(* IEC 61131-3 sources: plc-st-coding-agent/progress/evidence/f14_v3_parallel_20261112/jobs/custom_minimax-m27, 122 files *)

(* ---- public-easy-01.candidate_01.st ---- *)
FUNCTION_BLOCK FillingLineControl
VAR_INPUT
    bottleSensor         : BOOL;
    cleaningConfirmButton : BOOL;
    fillingConfirmButton  : BOOL;
    cappingConfirmButton  : BOOL;
    packingConfirmButton  : BOOL;
    finishedButton        : BOOL;
END_VAR

VAR_OUTPUT
    Pump_Motor      : BOOL;
    Filling_Valve   : BOOL;
    Capping_Machine : BOOL;
    Packing_Machine : BOOL;
    Completion_Light : BOOL;
END_VAR

VAR
    state : INT;
END_VAR

// State definitions:
// 0 = IDLE
// 1 = CLEANING
// 2 = FILLING
// 3 = CAPPING
// 4 = PACKAGING
// 5 = COMPLETED

// Reset all outputs at the start of each cycle
Pump_Motor      := FALSE;
Filling_Valve   := FALSE;
Capping_Machine := FALSE;
Packing_Machine := FALSE;
Completion_Light := FALSE;

CASE state OF
    0: // IDLE - Waiting for bottle
        IF bottleSensor THEN
            state := 1;
        END_IF;

    1: // CLEANING - Pump motor active
        Pump_Motor := TRUE;
        IF cleaningConfirmButton THEN
            state := 2;
        END_IF;

    2: // FILLING - Filling valve active
        Filling_Valve := TRUE;
        IF fillingConfirmButton THEN
            state := 3;
        END_IF;

    3: // CAPPING - Capping machine active
        Capping_Machine := TRUE;
        IF cappingConfirmButton THEN
            state := 4;
        END_IF;

    4: // PACKAGING - Packing machine active
        Packing_Machine := TRUE;
        IF packingConfirmButton THEN
            state := 5;
        END_IF;

    5: // COMPLETED - Completion light active
        Completion_Light := TRUE;
        IF finishedButton THEN
            state := 0;
        END_IF;

END_CASE;

END_FUNCTION_BLOCK

(* ---- public-easy-01.candidate_02.st ---- *)
FUNCTION_BLOCK FillingLineControl
VAR_INPUT
    bottleSensor          : BOOL;
    cleaningConfirmButton : BOOL;
    fillingConfirmButton  : BOOL;
    cappingConfirmButton  : BOOL;
    packingConfirmButton  : BOOL;
    finishedButton        : BOOL;
END_VAR

VAR_OUTPUT
    Pump_Motor       : BOOL;
    Filling_Valve    : BOOL;
    Capping_Machine  : BOOL;
    Packing_Machine  : BOOL;
    Completion_Light : BOOL;
END_VAR

VAR
    state : INT := 0;
END_VAR

// State: 0=IDLE, 1=CLEANING, 2=FILLING, 3=CAPPING, 4=PACKAGING, 5=COMPLETED

CASE state OF
    0: // IDLE
        IF bottleSensor THEN
            state := 1;
        END_IF;

    1: // CLEANING
        Pump_Motor := TRUE;
        IF cleaningConfirmButton THEN
            state := 2;
        END_IF;

    2: // FILLING
        Filling_Valve := TRUE;
        IF fillingConfirmButton THEN
            state := 3;
        END_IF;

    3: // CAPPING
        Capping_Machine := TRUE;
        IF cappingConfirmButton THEN
            state := 4;
        END_IF;

    4: // PACKAGING
        Packing_Machine := TRUE;
        IF packingConfirmButton THEN
            state := 5;
        END_IF;

    5: // COMPLETED
        Completion_Light := TRUE;
        IF finishedButton THEN
            state := 0;
        END_IF;

END_CASE;

END_FUNCTION_BLOCK

(* ---- public-easy-01.raw_candidate_01.st ---- *)
FUNCTION_BLOCK FillingLineControl
VAR_INPUT
    bottleSensor         : BOOL;
    cleaningConfirmButton : BOOL;
    fillingConfirmButton  : BOOL;
    cappingConfirmButton  : BOOL;
    packingConfirmButton  : BOOL;
    finishedButton        : BOOL;
END_VAR

VAR_OUTPUT
    Pump_Motor      : BOOL;
    Filling_Valve   : BOOL;
    Capping_Machine : BOOL;
    Packing_Machine : BOOL;
    Completion_Light : BOOL;
END_VAR

VAR
    state : INT;
END_VAR

// State definitions:
// 0 = IDLE
// 1 = CLEANING
// 2 = FILLING
// 3 = CAPPING
// 4 = PACKAGING
// 5 = COMPLETED

// Reset all outputs at the start of each cycle
Pump_Motor      := FALSE;
Filling_Valve   := FALSE;
Capping_Machine := FALSE;
Packing_Machine := FALSE;
Completion_Light := FALSE;

CASE state OF
    0: // IDLE - Waiting for bottle
        IF bottleSensor THEN
            state := 1;
        END_IF;

    1: // CLEANING - Pump motor active
        Pump_Motor := TRUE;
        IF cleaningConfirmButton THEN
            state := 2;
        END_IF;

    2: // FILLING - Filling valve active
        Filling_Valve := TRUE;
        IF fillingConfirmButton THEN
            state := 3;
        END_IF;

    3: // CAPPING - Capping machine active
        Capping_Machine := TRUE;
        IF cappingConfirmButton THEN
            state := 4;
        END_IF;

    4: // PACKAGING - Packing machine active
        Packing_Machine := TRUE;
        IF packingConfirmButton THEN
            state := 5;
        END_IF;

    5: // COMPLETED - Completion light active
        Completion_Light := TRUE;
        IF finishedButton THEN
            state := 0;
        END_IF;

END_CASE;

END_FUNCTION_BLOCK

(* ---- public-easy-01.raw_candidate_02.st ---- *)
FUNCTION_BLOCK FillingLineControl
VAR_INPUT
    bottleSensor          : BOOL;
    cleaningConfirmButton : BOOL;
    fillingConfirmButton  : BOOL;
    cappingConfirmButton  : BOOL;
    packingConfirmButton  : BOOL;
    finishedButton        : BOOL;
END_VAR

VAR_OUTPUT
    Pump_Motor       : BOOL;
    Filling_Valve    : BOOL;
    Capping_Machine  : BOOL;
    Packing_Machine  : BOOL;
    Completion_Light : BOOL;
END_VAR

VAR
    state : INT := 0;
END_VAR

// State: 0=IDLE, 1=CLEANING, 2=FILLING, 3=CAPPING, 4=PACKAGING, 5=COMPLETED

CASE state OF
    0: // IDLE
        IF bottleSensor THEN
            state := 1;
        END_IF;

    1: // CLEANING
        Pump_Motor := TRUE;
        IF cleaningConfirmButton THEN
            state := 2;
        END_IF;

    2: // FILLING
        Filling_Valve := TRUE;
        IF fillingConfirmButton THEN
            state := 3;
        END_IF;

    3: // CAPPING
        Capping_Machine := TRUE;
        IF cappingConfirmButton THEN
            state := 4;
        END_IF;

    4: // PACKAGING
        Packing_Machine := TRUE;
        IF packingConfirmButton THEN
            state := 5;
        END_IF;

    5: // COMPLETED
        Completion_Light := TRUE;
        IF finishedButton THEN
            state := 0;
        END_IF;

END_CASE;

END_FUNCTION_BLOCK

(* ---- public-easy-02.candidate_01.st ---- *)
FUNCTION_BLOCK FB_DualWordEdgeDetection
VAR
    prevValue : DWORD;
END_VAR

VAR_OUTPUT
    hasChanged      : BOOL := FALSE;
    hasRisingEdges  : BOOL := FALSE;
    risingBits      : DWORD := 0;
    noOfRisingBits  : USINT := 0;
    hasFallingEdges : BOOL := FALSE;
    fallingBits     : DWORD := 0;
    noOfFallingBits : USINT := 0;
END_VAR

VAR
    i : USINT;
END_VAR

risingBits  := value AND NOT prevValue;
fallingBits := NOT value AND prevValue;
hasChanged      := (value <> prevValue);
hasRisingEdges  := (risingBits <> 0);
hasFallingEdges := (fallingBits <> 0);

noOfRisingBits  := 0;
noOfFallingBits := 0;

FOR i := 0 TO 31 DO
    IF (risingBits AND SHL(DWORD#1, i)) <> 0 THEN
        noOfRisingBits := noOfRisingBits + 1;
    END_IF;
    IF (fallingBits AND SHL(DWORD#1, i)) <> 0 THEN
        noOfFallingBits := noOfFallingBits + 1;
    END_IF;
END_FOR;

prevValue := value;
END_FUNCTION_BLOCK

(* ---- public-easy-02.raw_candidate_01.st ---- *)
FUNCTION_BLOCK FB_DualWordEdgeDetection
VAR
    prevValue : DWORD;
END_VAR

VAR_OUTPUT
    hasChanged      : BOOL := FALSE;
    hasRisingEdges  : BOOL := FALSE;
    risingBits      : DWORD := 0;
    noOfRisingBits  : USINT := 0;
    hasFallingEdges : BOOL := FALSE;
    fallingBits     : DWORD := 0;
    noOfFallingBits : USINT := 0;
END_VAR

VAR
    i : USINT;
END_VAR

risingBits  := value AND NOT prevValue;
fallingBits := NOT value AND prevValue;
hasChanged      := (value <> prevValue);
hasRisingEdges  := (risingBits <> 0);
hasFallingEdges := (fallingBits <> 0);

noOfRisingBits  := 0;
noOfFallingBits := 0;

FOR i := 0 TO 31 DO
    IF (risingBits AND SHL(DWORD#1, i)) <> 0 THEN
        noOfRisingBits := noOfRisingBits + 1;
    END_IF;
    IF (fallingBits AND SHL(DWORD#1, i)) <> 0 THEN
        noOfFallingBits := noOfFallingBits + 1;
    END_IF;
END_FOR;

prevValue := value;
END_FUNCTION_BLOCK

(* ---- public-easy-03.candidate_01.st ---- *)
FUNCTION_BLOCK AlarmHysteresis
VAR_INPUT
    Value      : REAL;
    hiLevel    : REAL;
    loLevel    : REAL;
    hystWindow : REAL;
END_VAR

VAR_OUTPUT
    hiAlarm : BOOL;
    loAlarm : BOOL;
    error   : BOOL;
    status  : WORD;
END_VAR

VAR
END_VAR

error  := FALSE;
status := 16#0000;

IF loLevel >= hiLevel THEN
    error  := TRUE;
    status := 16#8001;
    RETURN;
END_IF;

IF hystWindow >= (hiLevel - loLevel) THEN
    error  := TRUE;
    status := 16#8002;
    RETURN;
END_IF;

IF Value > hiLevel THEN
    hiAlarm := TRUE;
ELSIF Value < (hiLevel - hystWindow) THEN
    hiAlarm := FALSE;
END_IF;

IF Value < loLevel THEN
    loAlarm := TRUE;
ELSIF Value > (loLevel + hystWindow) THEN
    loAlarm := FALSE;
END_IF;

END_FUNCTION_BLOCK

(* ---- public-easy-03.raw_candidate_01.st ---- *)
FUNCTION_BLOCK AlarmHysteresis
VAR_INPUT
    Value      : REAL;
    hiLevel    : REAL;
    loLevel    : REAL;
    hystWindow : REAL;
END_VAR

VAR_OUTPUT
    hiAlarm : BOOL;
    loAlarm : BOOL;
    error   : BOOL;
    status  : WORD;
END_VAR

VAR
END_VAR

error  := FALSE;
status := 16#0000;

IF loLevel >= hiLevel THEN
    error  := TRUE;
    status := 16#8001;
    RETURN;
END_IF;

IF hystWindow >= (hiLevel - loLevel) THEN
    error  := TRUE;
    status := 16#8002;
    RETURN;
END_IF;

IF Value > hiLevel THEN
    hiAlarm := TRUE;
ELSIF Value < (hiLevel - hystWindow) THEN
    hiAlarm := FALSE;
END_IF;

IF Value < loLevel THEN
    loAlarm := TRUE;
ELSIF Value > (loLevel + hystWindow) THEN
    loAlarm := FALSE;
END_IF;

END_FUNCTION_BLOCK

(* ---- public-easy-04.candidate_01.st ---- *)
FUNCTION_BLOCK JamPumpControl
VAR
    ViscosityValid : BOOL := FALSE;
    DebounceAccum  : LTIME  := LTIME#0s;
    PrevViscosity  : BOOL := FALSE;
END_VAR
VAR_OUTPUT
    VFD_RUN          : BOOL := FALSE;
    PUMP_MAINT_DUE   : BOOL := FALSE;
    PUMP_RUNTIME_ACC : LTIME  := LTIME#0s;
END_VAR
VAR_INPUT
    VISCOSITY_OK    : BOOL;
    PASTE_E_STOP_NC : BOOL;
    DebounceTime    : TIME;
    CycleTime       : TIME;
END_VAR

    // Emergency stop priority: immediate disable and clear debounce state
    IF NOT PASTE_E_STOP_NC THEN
        VFD_RUN        := FALSE;
        ViscosityValid := FALSE;
        DebounceAccum  := LTIME#0s;
        PrevViscosity  := FALSE;
        RETURN;
    END_IF;

    // Viscosity debouncing
    IF NOT VISCOSITY_OK THEN
        // Signal dropped: invalidate immediately and reset
        ViscosityValid := FALSE;
        DebounceAccum  := LTIME#0s;
        PrevViscosity  := FALSE;
    ELSE
        // Detect rising edge on VISCOSITY_OK
        IF NOT PrevViscosity THEN
            DebounceAccum := LTIME#0s;
        END_IF;

        // Accumulate debounce time for this cycle
        DebounceAccum := DebounceAccum + CycleTime;

        // Check if debounce threshold reached
        IF DebounceAccum >= DebounceTime THEN
            ViscosityValid := TRUE;
        END_IF;

        PrevViscosity := TRUE;
    END_IF;

    // Run permissive: E-stop OK AND viscosity condition valid AND signal present
    IF PASTE_E_STOP_NC AND ViscosityValid AND VISCOSITY_OK THEN
        VFD_RUN := TRUE;
    ELSE
        VFD_RUN := FALSE;
    END_IF;

    // Accumulate runtime only while pump is running
    IF VFD_RUN THEN
        PUMP_RUNTIME_ACC := PUMP_RUNTIME_ACC + CycleTime;
    END_IF;

    // Maintenance indication at 500 hours (informational, non-blocking)
    IF PUMP_RUNTIME_ACC >= T#500h THEN
        PUMP_MAINT_DUE := TRUE;
    END_IF;

END_FUNCTION_BLOCK

(* ---- public-easy-04.candidate_02.st ---- *)
FUNCTION_BLOCK JamPumpControl
VAR
    ViscosityValid : BOOL := FALSE;
    DebounceAccum  : LTIME  := LTIME#0s;
    PrevViscosity  : BOOL := FALSE;
END_VAR
VAR_OUTPUT
    VFD_RUN          : BOOL := FALSE;
    PUMP_MAINT_DUE   : BOOL := FALSE;
    PUMP_RUNTIME_ACC : LTIME  := LTIME#0s;
END_VAR
VAR_INPUT
    VISCOSITY_OK    : BOOL;
    PASTE_E_STOP_NC : BOOL;
    DebounceTime    : TIME;
    CycleTime       : TIME;
END_VAR
    // Emergency stop priority: immediate disable and clear debounce state
    IF NOT PASTE_E_STOP_NC THEN
        VFD_RUN        := FALSE;
        ViscosityValid := FALSE;
        DebounceAccum  := LTIME#0s;
        PrevViscosity  := FALSE;
        RETURN;
    END_IF;

    // Viscosity debouncing
    IF NOT VISCOSITY_OK THEN
        ViscosityValid := FALSE;
        DebounceAccum  := LTIME#0s;
        PrevViscosity  := FALSE;
    ELSE
        IF NOT PrevViscosity THEN
            DebounceAccum := LTIME#0s;
        END_IF;

        DebounceAccum := DebounceAccum + TO_LTIME(TO_ULINT(CycleTime));

        IF DebounceAccum >= TO_LTIME(TO_ULINT(DebounceTime)) THEN
            ViscosityValid := TRUE;
        END_IF;

        PrevViscosity := TRUE;
    END_IF;

    // Run permissive
    IF PASTE_E_STOP_NC AND ViscosityValid AND VISCOSITY_OK THEN
        VFD_RUN := TRUE;
    ELSE
        VFD_RUN := FALSE;
    END_IF;

    // Accumulate runtime only while pump is running
    IF VFD_RUN THEN
        PUMP_RUNTIME_ACC := PUMP_RUNTIME_ACC + TO_LTIME(TO_ULINT(CycleTime));
    END_IF;

    // Maintenance indication at 500 hours
    IF PUMP_RUNTIME_ACC >= LTIME#500h THEN
        PUMP_MAINT_DUE := TRUE;
    END_IF;

END_FUNCTION_BLOCK

(* ---- public-easy-04.raw_candidate_01.st ---- *)
FUNCTION_BLOCK JamPumpControl
VAR
    ViscosityValid : BOOL := FALSE;
    DebounceAccum  : LTIME  := LTIME#0s;
    PrevViscosity  : BOOL := FALSE;
END_VAR
VAR_OUTPUT
    VFD_RUN          : BOOL := FALSE;
    PUMP_MAINT_DUE   : BOOL := FALSE;
    PUMP_RUNTIME_ACC : LTIME  := LTIME#0s;
END_VAR
VAR_INPUT
    VISCOSITY_OK    : BOOL;
    PASTE_E_STOP_NC : BOOL;
    DebounceTime    : TIME;
    CycleTime       : TIME;
END_VAR

    // Emergency stop priority: immediate disable and clear debounce state
    IF NOT PASTE_E_STOP_NC THEN
        VFD_RUN        := FALSE;
        ViscosityValid := FALSE;
        DebounceAccum  := LTIME#0s;
        PrevViscosity  := FALSE;
        RETURN;
    END_IF;

    // Viscosity debouncing
    IF NOT VISCOSITY_OK THEN
        // Signal dropped: invalidate immediately and reset
        ViscosityValid := FALSE;
        DebounceAccum  := LTIME#0s;
        PrevViscosity  := FALSE;
    ELSE
        // Detect rising edge on VISCOSITY_OK
        IF NOT PrevViscosity THEN
            DebounceAccum := LTIME#0s;
        END_IF;

        // Accumulate debounce time for this cycle
        DebounceAccum := DebounceAccum + CycleTime;

        // Check if debounce threshold reached
        IF DebounceAccum >= DebounceTime THEN
            ViscosityValid := TRUE;
        END_IF;

        PrevViscosity := TRUE;
    END_IF;

    // Run permissive: E-stop OK AND viscosity condition valid AND signal present
    IF PASTE_E_STOP_NC AND ViscosityValid AND VISCOSITY_OK THEN
        VFD_RUN := TRUE;
    ELSE
        VFD_RUN := FALSE;
    END_IF;

    // Accumulate runtime only while pump is running
    IF VFD_RUN THEN
        PUMP_RUNTIME_ACC := PUMP_RUNTIME_ACC + CycleTime;
    END_IF;

    // Maintenance indication at 500 hours (informational, non-blocking)
    IF PUMP_RUNTIME_ACC >= T#500h THEN
        PUMP_MAINT_DUE := TRUE;
    END_IF;

END_FUNCTION_BLOCK

(* ---- public-easy-04.raw_candidate_02.st ---- *)
FUNCTION_BLOCK JamPumpControl
VAR
    ViscosityValid : BOOL := FALSE;
    DebounceAccum  : LTIME  := LTIME#0s;
    PrevViscosity  : BOOL := FALSE;
END_VAR
VAR_OUTPUT
    VFD_RUN          : BOOL := FALSE;
    PUMP_MAINT_DUE   : BOOL := FALSE;
    PUMP_RUNTIME_ACC : LTIME  := LTIME#0s;
END_VAR
VAR_INPUT
    VISCOSITY_OK    : BOOL;
    PASTE_E_STOP_NC : BOOL;
    DebounceTime    : TIME;
    CycleTime       : TIME;
END_VAR
    // Emergency stop priority: immediate disable and clear debounce state
    IF NOT PASTE_E_STOP_NC THEN
        VFD_RUN        := FALSE;
        ViscosityValid := FALSE;
        DebounceAccum  := LTIME#0s;
        PrevViscosity  := FALSE;
        RETURN;
    END_IF;

    // Viscosity debouncing
    IF NOT VISCOSITY_OK THEN
        ViscosityValid := FALSE;
        DebounceAccum  := LTIME#0s;
        PrevViscosity  := FALSE;
    ELSE
        IF NOT PrevViscosity THEN
            DebounceAccum := LTIME#0s;
        END_IF;

        DebounceAccum := DebounceAccum + TO_LTIME(TO_ULINT(CycleTime));

        IF DebounceAccum >= TO_LTIME(TO_ULINT(DebounceTime)) THEN
            ViscosityValid := TRUE;
        END_IF;

        PrevViscosity := TRUE;
    END_IF;

    // Run permissive
    IF PASTE_E_STOP_NC AND ViscosityValid AND VISCOSITY_OK THEN
        VFD_RUN := TRUE;
    ELSE
        VFD_RUN := FALSE;
    END_IF;

    // Accumulate runtime only while pump is running
    IF VFD_RUN THEN
        PUMP_RUNTIME_ACC := PUMP_RUNTIME_ACC + TO_LTIME(TO_ULINT(CycleTime));
    END_IF;

    // Maintenance indication at 500 hours
    IF PUMP_RUNTIME_ACC >= LTIME#500h THEN
        PUMP_MAINT_DUE := TRUE;
    END_IF;

END_FUNCTION_BLOCK

(* ---- public-easy-05.candidate_01.st ---- *)
FUNCTION_BLOCK Weld_Gap_Alarm
VAR_INPUT
    Gap_Exceeded    : BOOL;
    Weld_E_Stop_NC  : BOOL;
    DebounceTime    : TIME;
END_VAR
VAR_OUTPUT
    Operator_Alert        : BOOL := FALSE;
    Weld_Soft_Start_Active: BOOL := FALSE;
END_VAR
VAR
    State           : (EStop, Init, Monitor) := Init;
    Init_Timer      : TON;
    Gap_Debounce    : TON;
    Gap_Debounced   : BOOL := FALSE;
    Gap_Accumulated : LTIME := LTIME#0s;
    CycleCount      : UINT := 0;
END_VAR

// EStop has highest priority - immediate reaction before any other logic
IF NOT Weld_E_Stop_NC THEN
    Operator_Alert := FALSE;
    Weld_Soft_Start_Active := FALSE;
    Gap_Debounced := FALSE;
    Gap_Accumulated := LTIME#0s;
    Gap_Debounce(IN := FALSE);
    Gap_Debounce.PT := T#0ms;
    Init_Timer(IN := FALSE);
    Init_Timer.PT := T#0ms;
    Init_Timer.Q := FALSE;
    State := EStop;
    RETURN;
END_IF;

// EStop released - restart initialization timer
IF State = EStop THEN
    State := Init;
    Init_Timer(IN := FALSE);
END_IF;

// State machine for initialization and monitoring
CASE State OF
    Init:
        // Begin 5-second initialization inhibition
        Init_Timer(IN := TRUE, PT := T#5s);
        Weld_Soft_Start_Active := TRUE;
        Operator_Alert := FALSE;
        Gap_Debounced := FALSE;
        Gap_Accumulated := LTIME#0s;
        Gap_Debounce(IN := FALSE);
        Gap_Debounce.PT := T#0ms;

        // Transition to monitoring after initialization completes
        IF Init_Timer.Q THEN
            State := Monitor;
            Weld_Soft_Start_Active := FALSE;
        END_IF;

    Monitor:
        Init_Timer(IN := FALSE);
        Init_Timer.Q := FALSE;
        Weld_Soft_Start_Active := FALSE;

        // Gap monitoring with debounce
        IF Gap_Exceeded THEN
            // Accumulate debounce time using cycle-based increment
            Gap_Accumulated := Gap_Accumulated + TO_LTIME(CycleCount);

            // Check if debounce threshold reached
            IF Gap_Accumulated >= TO_LTIME(DebounceTime) THEN
                Gap_Debounced := TRUE;
                Operator_Alert := TRUE;
            END_IF;
        ELSE
            // Signal is FALSE - clear alarm and reset debounce
            Gap_Debounced := FALSE;
            Operator_Alert := FALSE;
            Gap_Accumulated := LTIME#0s;
        END_IF;
END_CASE;

// Track cycle time for debounce accumulation
CycleCount := TO_UINT(T#1ms) / TO_UINT(T#1ms);

END_FUNCTION_BLOCK

(* ---- public-easy-05.candidate_02.st ---- *)
TYPE GapAlarmState :
(
    EStop  := 0,
    Init   := 1,
    Monitor := 2
) END_TYPE;

FUNCTION_BLOCK Weld_Gap_Alarm
VAR_INPUT
    Gap_Exceeded   : BOOL;
    Weld_E_Stop_NC : BOOL;
    DebounceTime   : TIME;
END_VAR
VAR_OUTPUT
    Operator_Alert        : BOOL := FALSE;
    Weld_Soft_Start_Active: BOOL := FALSE;
END_VAR
VAR
    State        : GapAlarmState := Init;
    Init_Timer   : TON;
    Gap_Debounce : TON;
END_VAR

// EStop has highest priority
IF NOT Weld_E_Stop_NC THEN
    Operator_Alert        := FALSE;
    Weld_Soft_Start_Active := FALSE;
    Init_Timer(IN := FALSE);
    Gap_Debounce(IN := FALSE);
    State := EStop;
    RETURN;
END_IF;

// EStop released - transition to initialization
IF State = EStop THEN
    State := Init;
END_IF;

CASE State OF
    Init:
        Init_Timer(IN := TRUE, PT := T#5s);
        Weld_Soft_Start_Active := TRUE;
        Operator_Alert := FALSE;
        Gap_Debounce(IN := FALSE);

        IF Init_Timer.Q THEN
            State := Monitor;
            Weld_Soft_Start_Active := FALSE;
        END_IF;

    Monitor:
        Init_Timer(IN := FALSE);
        Weld_Soft_Start_Active := FALSE;

        // Debounce gap signal: timer accumulates while TRUE,
        // resets when FALSE (ET tracks elapsed time)
        Gap_Debounce(IN := Gap_Exceeded, PT := DebounceTime);

        IF Gap_Debounce.Q THEN
            Operator_Alert := TRUE;
        ELSE
            Operator_Alert := FALSE;
        END_IF;
END_CASE;

END_FUNCTION_BLOCK

(* ---- public-easy-05.raw_candidate_01.st ---- *)
FUNCTION_BLOCK Weld_Gap_Alarm
VAR_INPUT
    Gap_Exceeded    : BOOL;
    Weld_E_Stop_NC  : BOOL;
    DebounceTime    : TIME;
END_VAR
VAR_OUTPUT
    Operator_Alert        : BOOL := FALSE;
    Weld_Soft_Start_Active: BOOL := FALSE;
END_VAR
VAR
    State           : (EStop, Init, Monitor) := Init;
    Init_Timer      : TON;
    Gap_Debounce    : TON;
    Gap_Debounced   : BOOL := FALSE;
    Gap_Accumulated : LTIME := LTIME#0s;
    CycleCount      : UINT := 0;
END_VAR

// EStop has highest priority - immediate reaction before any other logic
IF NOT Weld_E_Stop_NC THEN
    Operator_Alert := FALSE;
    Weld_Soft_Start_Active := FALSE;
    Gap_Debounced := FALSE;
    Gap_Accumulated := LTIME#0s;
    Gap_Debounce(IN := FALSE);
    Gap_Debounce.PT := T#0ms;
    Init_Timer(IN := FALSE);
    Init_Timer.PT := T#0ms;
    Init_Timer.Q := FALSE;
    State := EStop;
    RETURN;
END_IF;

// EStop released - restart initialization timer
IF State = EStop THEN
    State := Init;
    Init_Timer(IN := FALSE);
END_IF;

// State machine for initialization and monitoring
CASE State OF
    Init:
        // Begin 5-second initialization inhibition
        Init_Timer(IN := TRUE, PT := T#5s);
        Weld_Soft_Start_Active := TRUE;
        Operator_Alert := FALSE;
        Gap_Debounced := FALSE;
        Gap_Accumulated := LTIME#0s;
        Gap_Debounce(IN := FALSE);
        Gap_Debounce.PT := T#0ms;

        // Transition to monitoring after initialization completes
        IF Init_Timer.Q THEN
            State := Monitor;
            Weld_Soft_Start_Active := FALSE;
        END_IF;

    Monitor:
        Init_Timer(IN := FALSE);
        Init_Timer.Q := FALSE;
        Weld_Soft_Start_Active := FALSE;

        // Gap monitoring with debounce
        IF Gap_Exceeded THEN
            // Accumulate debounce time using cycle-based increment
            Gap_Accumulated := Gap_Accumulated + TO_LTIME(CycleCount);

            // Check if debounce threshold reached
            IF Gap_Accumulated >= TO_LTIME(DebounceTime) THEN
                Gap_Debounced := TRUE;
                Operator_Alert := TRUE;
            END_IF;
        ELSE
            // Signal is FALSE - clear alarm and reset debounce
            Gap_Debounced := FALSE;
            Operator_Alert := FALSE;
            Gap_Accumulated := LTIME#0s;
        END_IF;
END_CASE;

// Track cycle time for debounce accumulation
CycleCount := TO_UINT(T#1ms) / TO_UINT(T#1ms);

END_FUNCTION_BLOCK

(* ---- public-easy-05.raw_candidate_02.st ---- *)
TYPE GapAlarmState :
(
    EStop  := 0,
    Init   := 1,
    Monitor := 2
) END_TYPE

FUNCTION_BLOCK Weld_Gap_Alarm
VAR_INPUT
    Gap_Exceeded   : BOOL;
    Weld_E_Stop_NC : BOOL;
    DebounceTime   : TIME;
END_VAR
VAR_OUTPUT
    Operator_Alert        : BOOL := FALSE;
    Weld_Soft_Start_Active: BOOL := FALSE;
END_VAR
VAR
    State        : GapAlarmState := Init;
    Init_Timer   : TON;
    Gap_Debounce : TON;
END_VAR

// EStop has highest priority
IF NOT Weld_E_Stop_NC THEN
    Operator_Alert        := FALSE;
    Weld_Soft_Start_Active := FALSE;
    Init_Timer(IN := FALSE);
    Gap_Debounce(IN := FALSE);
    State := EStop;
    RETURN;
END_IF;

// EStop released - transition to initialization
IF State = EStop THEN
    State := Init;
END_IF;

CASE State OF
    Init:
        Init_Timer(IN := TRUE, PT := T#5s);
        Weld_Soft_Start_Active := TRUE;
        Operator_Alert := FALSE;
        Gap_Debounce(IN := FALSE);

        IF Init_Timer.Q THEN
            State := Monitor;
            Weld_Soft_Start_Active := FALSE;
        END_IF;

    Monitor:
        Init_Timer(IN := FALSE);
        Weld_Soft_Start_Active := FALSE;

        // Debounce gap signal: timer accumulates while TRUE,
        // resets when FALSE (ET tracks elapsed time)
        Gap_Debounce(IN := Gap_Exceeded, PT := DebounceTime);

        IF Gap_Debounce.Q THEN
            Operator_Alert := TRUE;
        ELSE
            Operator_Alert := FALSE;
        END_IF;
END_CASE;

END_FUNCTION_BLOCK

(* ---- public-easy-06.candidate_01.st ---- *)
FUNCTION_BLOCK AerationBlowerControl
VAR_INPUT
    DO_LOW : BOOL;
    AERATION_E_STOP_NC : BOOL;
END_VAR

VAR_OUTPUT
    BLOWER_RUN : BOOL := FALSE;
    AERATION_BLOWER_CYCLE_COUNT : UINT := 0;
END_VAR

VAR
    StartDelayTimer : TON;
    BlowerRunPrev : BOOL := FALSE;
END_VAR

    // Start delay timing when both DO_LOW and E-stop inactive (NC = TRUE)
    IF DO_LOW AND AERATION_E_STOP_NC THEN
        // Start the 5-second timer
        StartDelayTimer(IN := TRUE, PT := T#5S);

        // BLOWER_RUN only TRUE after timer completes
        IF StartDelayTimer.Q THEN
            BLOWER_RUN := TRUE;
        ELSE
            BLOWER_RUN := FALSE;
        END_IF;
    ELSE
        // Conditions lost: reset timer and disable blower
        StartDelayTimer(IN := FALSE);
        BLOWER_RUN := FALSE;
    END_IF;

    // Count FALSE-to-TRUE transitions of BLOWER_RUN
    IF BLOWER_RUN AND NOT BlowerRunPrev THEN
        AERATION_BLOWER_CYCLE_COUNT := AERATION_BLOWER_CYCLE_COUNT + 1;
    END_IF;

    // Store previous state for edge detection
    BlowerRunPrev := BLOWER_RUN;

END_FUNCTION_BLOCK

(* ---- public-easy-06.raw_candidate_01.st ---- *)
FUNCTION_BLOCK AerationBlowerControl
VAR_INPUT
    DO_LOW : BOOL;
    AERATION_E_STOP_NC : BOOL;
END_VAR

VAR_OUTPUT
    BLOWER_RUN : BOOL := FALSE;
    AERATION_BLOWER_CYCLE_COUNT : UINT := 0;
END_VAR

VAR
    StartDelayTimer : TON;
    BlowerRunPrev : BOOL := FALSE;
END_VAR

    // Start delay timing when both DO_LOW and E-stop inactive (NC = TRUE)
    IF DO_LOW AND AERATION_E_STOP_NC THEN
        // Start the 5-second timer
        StartDelayTimer(IN := TRUE, PT := T#5S);

        // BLOWER_RUN only TRUE after timer completes
        IF StartDelayTimer.Q THEN
            BLOWER_RUN := TRUE;
        ELSE
            BLOWER_RUN := FALSE;
        END_IF;
    ELSE
        // Conditions lost: reset timer and disable blower
        StartDelayTimer(IN := FALSE);
        BLOWER_RUN := FALSE;
    END_IF;

    // Count FALSE-to-TRUE transitions of BLOWER_RUN
    IF BLOWER_RUN AND NOT BlowerRunPrev THEN
        AERATION_BLOWER_CYCLE_COUNT := AERATION_BLOWER_CYCLE_COUNT + 1;
    END_IF;

    // Store previous state for edge detection
    BlowerRunPrev := BLOWER_RUN;

END_FUNCTION_BLOCK

(* ---- public-hard-01.candidate_01.st ---- *)
FUNCTION_BLOCK MaterialProportioningControl
VAR_INPUT
    estop            : BOOL;
    opeMode          : BOOL;
    valveAStart      : BOOL;
    valveBStart      : BOOL;
    valveCStart      : BOOL;
    valveDStart      : BOOL;
    mixMotorStart    : BOOL;
    autoStart        : BOOL;
    processMode      : BOOL;
    levelSensor      : INT;
    mixMotorComplete : BOOL;
END_VAR
VAR_OUTPUT
    valveARun    : BOOL;
    valveBRun    : BOOL;
    valveCRun    : BOOL;
    valveDRun    : BOOL;
    mixMotorRun  : BOOL;
END_VAR
VAR
    State          : INT;
    StateNext      : INT;
    autoStarted    : BOOL;
    valveAToggled  : BOOL;
    valveBToggled  : BOOL;
    valveCToggled  : BOOL;
    valveDToggled  : BOOL;
    motorToggled   : BOOL;
    lastAutoStart  : BOOL;
    lastValveAStart : BOOL;
    lastValveBStart : BOOL;
    lastValveCStart : BOOL;
    lastValveDStart : BOOL;
    lastMixMotorStart : BOOL;
END_VAR

VAR CONSTANT
    AUTO_IDLE       : INT := 0;
    AUTO_FILL_A     : INT := 1;
    AUTO_FILL_B     : INT := 2;
    AUTO_FILL_C     : INT := 3;
    AUTO_MIXING     : INT := 4;
    AUTO_DRAIN      : INT := 5;
END_VAR

    lastAutoStart := autoStart;
    lastValveAStart := valveAStart;
    lastValveBStart := valveBStart;
    lastValveCStart := valveCStart;
    lastValveDStart := valveDStart;
    lastMixMotorStart := mixMotorStart;

    valveARun := FALSE;
    valveBRun := FALSE;
    valveCRun := FALSE;
    valveDRun := FALSE;
    mixMotorRun := FALSE;

    IF NOT estop THEN
        State := AUTO_IDLE;
        autoStarted := FALSE;
        valveAToggled := FALSE;
        valveBToggled := FALSE;
        valveCToggled := FALSE;
        valveDToggled := FALSE;
        motorToggled := FALSE;
        RETURN;
    END_IF;

    IF NOT opeMode THEN
        State := AUTO_IDLE;
        autoStarted := FALSE;

        IF valveAStart AND NOT lastValveAStart THEN
            valveAToggled := NOT valveAToggled;
        END_IF;

        IF valveBStart AND NOT lastValveBStart THEN
            valveBToggled := NOT valveBToggled;
        END_IF;

        IF valveCStart AND NOT lastValveCStart THEN
            valveCToggled := NOT valveCToggled;
        END_IF;

        IF valveDStart AND NOT lastValveDStart THEN
            valveDToggled := NOT valveDToggled;
        END_IF;

        IF mixMotorStart AND NOT lastMixMotorStart THEN
            motorToggled := NOT motorToggled;
        END_IF;

        valveARun := valveAToggled;
        valveBRun := valveBToggled;
        valveCRun := valveCToggled;
        valveDRun := valveDToggled;
        mixMotorRun := motorToggled;

        RETURN;
    END_IF;

    CASE State OF
        AUTO_IDLE:
            autoStarted := FALSE;
            valveAToggled := FALSE;
            valveBToggled := FALSE;
            valveCToggled := FALSE;
            valveDToggled := FALSE;
            motorToggled := FALSE;
            IF autoStart AND NOT lastAutoStart THEN
                State := AUTO_FILL_A;
            END_IF;

        AUTO_FILL_A:
            valveARun := TRUE;
            IF levelSensor >= 50 THEN
                valveARun := FALSE;
                State := AUTO_FILL_B;
            END_IF;

        AUTO_FILL_B:
            valveBRun := TRUE;
            IF levelSensor >= 80 THEN
                valveBRun := FALSE;
                IF NOT processMode THEN
                    State := AUTO_MIXING;
                ELSE
                    State := AUTO_FILL_C;
                END_IF;
            END_IF;

        AUTO_FILL_C:
            valveCRun := TRUE;
            IF levelSensor >= 100 THEN
                valveCRun := FALSE;
                State := AUTO_MIXING;
            END_IF;

        AUTO_MIXING:
            mixMotorRun := TRUE;
            IF mixMotorComplete THEN
                mixMotorRun := FALSE;
                State := AUTO_DRAIN;
            END_IF;

        AUTO_DRAIN:
            valveDRun := TRUE;

    END_CASE;

END_FUNCTION_BLOCK

(* ---- public-hard-01.candidate_02.st ---- *)
FUNCTION_BLOCK MaterialProportioningControl
VAR_INPUT
    estop            : BOOL;
    opeMode          : BOOL;
    valveAStart      : BOOL;
    valveBStart      : BOOL;
    valveCStart      : BOOL;
    valveDStart      : BOOL;
    mixMotorStart    : BOOL;
    autoStart        : BOOL;
    processMode      : BOOL;
    levelSensor      : INT;
    mixMotorComplete : BOOL;
END_VAR
VAR_OUTPUT
    valveARun    : BOOL;
    valveBRun    : BOOL;
    valveCRun    : BOOL;
    valveDRun    : BOOL;
    mixMotorRun  : BOOL;
END_VAR
VAR
    State             : INT;
    valveAToggled     : BOOL;
    valveBToggled     : BOOL;
    valveCToggled     : BOOL;
    valveDToggled     : BOOL;
    motorToggled      : BOOL;
    prevAutoStart     : BOOL;
    prevValveAStart   : BOOL;
    prevValveBStart   : BOOL;
    prevValveCStart   : BOOL;
    prevValveDStart   : BOOL;
    prevMixMotorStart : BOOL;
END_VAR

VAR CONSTANT
    AUTO_IDLE   : INT := 0;
    AUTO_FILL_A : INT := 1;
    AUTO_FILL_B : INT := 2;
    AUTO_FILL_C : INT := 3;
    AUTO_MIXING : INT := 4;
    AUTO_DRAIN  : INT := 5;
END_VAR

    valveARun := FALSE;
    valveBRun := FALSE;
    valveCRun := FALSE;
    valveDRun := FALSE;
    mixMotorRun := FALSE;

    IF NOT estop THEN
        State := AUTO_IDLE;
        valveAToggled := FALSE;
        valveBToggled := FALSE;
        valveCToggled := FALSE;
        valveDToggled := FALSE;
        motorToggled := FALSE;
        prevAutoStart := FALSE;
        prevValveAStart := FALSE;
        prevValveBStart := FALSE;
        prevValveCStart := FALSE;
        prevValveDStart := FALSE;
        prevMixMotorStart := FALSE;
        RETURN;
    END_IF;

    IF NOT opeMode THEN
        State := AUTO_IDLE;

        IF valveAStart AND NOT prevValveAStart THEN
            valveAToggled := NOT valveAToggled;
        END_IF;
        IF valveBStart AND NOT prevValveBStart THEN
            valveBToggled := NOT valveBToggled;
        END_IF;
        IF valveCStart AND NOT prevValveCStart THEN
            valveCToggled := NOT valveCToggled;
        END_IF;
        IF valveDStart AND NOT prevValveDStart THEN
            valveDToggled := NOT valveDToggled;
        END_IF;
        IF mixMotorStart AND NOT prevMixMotorStart THEN
            motorToggled := NOT motorToggled;
        END_IF;

        valveARun := valveAToggled;
        valveBRun := valveBToggled;
        valveCRun := valveCToggled;
        valveDRun := valveDToggled;
        mixMotorRun := motorToggled;
    ELSE
        CASE State OF
            AUTO_IDLE:
                valveAToggled := FALSE;
                valveBToggled := FALSE;
                valveCToggled := FALSE;
                valveDToggled := FALSE;
                motorToggled := FALSE;
                IF autoStart AND NOT prevAutoStart THEN
                    State := AUTO_FILL_A;
                END_IF;

            AUTO_FILL_A:
                valveARun := TRUE;
                IF levelSensor >= 50 THEN
                    valveARun := FALSE;
                    State := AUTO_FILL_B;
                END_IF;

            AUTO_FILL_B:
                valveBRun := TRUE;
                IF levelSensor >= 80 THEN
                    valveBRun := FALSE;
                    IF NOT processMode THEN
                        State := AUTO_MIXING;
                    ELSE
                        State := AUTO_FILL_C;
                    END_IF;
                END_IF;

            AUTO_FILL_C:
                valveCRun := TRUE;
                IF levelSensor >= 100 THEN
                    valveCRun := FALSE;
                    State := AUTO_MIXING;
                END_IF;

            AUTO_MIXING:
                mixMotorRun := TRUE;
                IF mixMotorComplete THEN
                    mixMotorRun := FALSE;
                    State := AUTO_DRAIN;
                END_IF;

            AUTO_DRAIN:
                valveDRun := TRUE;
        END_CASE;
    END_IF;

    prevAutoStart := autoStart;
    prevValveAStart := valveAStart;
    prevValveBStart := valveBStart;
    prevValveCStart := valveCStart;
    prevValveDStart := valveDStart;
    prevMixMotorStart := mixMotorStart;

END_FUNCTION_BLOCK

(* ---- public-hard-01.raw_candidate_01.st ---- *)
FUNCTION_BLOCK MaterialProportioningControl
VAR_INPUT
    estop            : BOOL;
    opeMode          : BOOL;
    valveAStart      : BOOL;
    valveBStart      : BOOL;
    valveCStart      : BOOL;
    valveDStart      : BOOL;
    mixMotorStart    : BOOL;
    autoStart        : BOOL;
    processMode      : BOOL;
    levelSensor      : INT;
    mixMotorComplete : BOOL;
END_VAR
VAR_OUTPUT
    valveARun    : BOOL;
    valveBRun    : BOOL;
    valveCRun    : BOOL;
    valveDRun    : BOOL;
    mixMotorRun  : BOOL;
END_VAR
VAR
    State          : INT;
    StateNext      : INT;
    autoStarted    : BOOL;
    valveAToggled  : BOOL;
    valveBToggled  : BOOL;
    valveCToggled  : BOOL;
    valveDToggled  : BOOL;
    motorToggled   : BOOL;
    lastAutoStart  : BOOL;
    lastValveAStart : BOOL;
    lastValveBStart : BOOL;
    lastValveCStart : BOOL;
    lastValveDStart : BOOL;
    lastMixMotorStart : BOOL;
END_VAR

VAR CONSTANT
    AUTO_IDLE       : INT := 0;
    AUTO_FILL_A     : INT := 1;
    AUTO_FILL_B     : INT := 2;
    AUTO_FILL_C     : INT := 3;
    AUTO_MIXING     : INT := 4;
    AUTO_DRAIN      : INT := 5;
END_VAR

    lastAutoStart := autoStart;
    lastValveAStart := valveAStart;
    lastValveBStart := valveBStart;
    lastValveCStart := valveCStart;
    lastValveDStart := valveDStart;
    lastMixMotorStart := mixMotorStart;

    valveARun := FALSE;
    valveBRun := FALSE;
    valveCRun := FALSE;
    valveDRun := FALSE;
    mixMotorRun := FALSE;

    IF NOT estop THEN
        State := AUTO_IDLE;
        autoStarted := FALSE;
        valveAToggled := FALSE;
        valveBToggled := FALSE;
        valveCToggled := FALSE;
        valveDToggled := FALSE;
        motorToggled := FALSE;
        RETURN;
    END_IF

    IF NOT opeMode THEN
        State := AUTO_IDLE;
        autoStarted := FALSE;

        IF valveAStart AND NOT lastValveAStart THEN
            valveAToggled := NOT valveAToggled;
        END_IF

        IF valveBStart AND NOT lastValveBStart THEN
            valveBToggled := NOT valveBToggled;
        END_IF

        IF valveCStart AND NOT lastValveCStart THEN
            valveCToggled := NOT valveCToggled;
        END_IF

        IF valveDStart AND NOT lastValveDStart THEN
            valveDToggled := NOT valveDToggled;
        END_IF

        IF mixMotorStart AND NOT lastMixMotorStart THEN
            motorToggled := NOT motorToggled;
        END_IF

        valveARun := valveAToggled;
        valveBRun := valveBToggled;
        valveCRun := valveCToggled;
        valveDRun := valveDToggled;
        mixMotorRun := motorToggled;

        RETURN;
    END_IF

    CASE State OF
        AUTO_IDLE:
            autoStarted := FALSE;
            valveAToggled := FALSE;
            valveBToggled := FALSE;
            valveCToggled := FALSE;
            valveDToggled := FALSE;
            motorToggled := FALSE;
            IF autoStart AND NOT lastAutoStart THEN
                State := AUTO_FILL_A;
            END_IF;

        AUTO_FILL_A:
            valveARun := TRUE;
            IF levelSensor >= 50 THEN
                valveARun := FALSE;
                State := AUTO_FILL_B;
            END_IF;

        AUTO_FILL_B:
            valveBRun := TRUE;
            IF levelSensor >= 80 THEN
                valveBRun := FALSE;
                IF NOT processMode THEN
                    State := AUTO_MIXING;
                ELSE
                    State := AUTO_FILL_C;
                END_IF;
            END_IF;

        AUTO_FILL_C:
            valveCRun := TRUE;
            IF levelSensor >= 100 THEN
                valveCRun := FALSE;
                State := AUTO_MIXING;
            END_IF;

        AUTO_MIXING:
            mixMotorRun := TRUE;
            IF mixMotorComplete THEN
                mixMotorRun := FALSE;
                State := AUTO_DRAIN;
            END_IF;

        AUTO_DRAIN:
            valveDRun := TRUE;

    END_CASE;

END_FUNCTION_BLOCK

(* ---- public-hard-01.raw_candidate_02.st ---- *)
FUNCTION_BLOCK MaterialProportioningControl
VAR_INPUT
    estop            : BOOL;
    opeMode          : BOOL;
    valveAStart      : BOOL;
    valveBStart      : BOOL;
    valveCStart      : BOOL;
    valveDStart      : BOOL;
    mixMotorStart    : BOOL;
    autoStart        : BOOL;
    processMode      : BOOL;
    levelSensor      : INT;
    mixMotorComplete : BOOL;
END_VAR
VAR_OUTPUT
    valveARun    : BOOL;
    valveBRun    : BOOL;
    valveCRun    : BOOL;
    valveDRun    : BOOL;
    mixMotorRun  : BOOL;
END_VAR
VAR
    State             : INT;
    valveAToggled     : BOOL;
    valveBToggled     : BOOL;
    valveCToggled     : BOOL;
    valveDToggled     : BOOL;
    motorToggled      : BOOL;
    prevAutoStart     : BOOL;
    prevValveAStart   : BOOL;
    prevValveBStart   : BOOL;
    prevValveCStart   : BOOL;
    prevValveDStart   : BOOL;
    prevMixMotorStart : BOOL;
END_VAR

VAR CONSTANT
    AUTO_IDLE   : INT := 0;
    AUTO_FILL_A : INT := 1;
    AUTO_FILL_B : INT := 2;
    AUTO_FILL_C : INT := 3;
    AUTO_MIXING : INT := 4;
    AUTO_DRAIN  : INT := 5;
END_VAR

    valveARun := FALSE;
    valveBRun := FALSE;
    valveCRun := FALSE;
    valveDRun := FALSE;
    mixMotorRun := FALSE;

    IF NOT estop THEN
        State := AUTO_IDLE;
        valveAToggled := FALSE;
        valveBToggled := FALSE;
        valveCToggled := FALSE;
        valveDToggled := FALSE;
        motorToggled := FALSE;
        prevAutoStart := FALSE;
        prevValveAStart := FALSE;
        prevValveBStart := FALSE;
        prevValveCStart := FALSE;
        prevValveDStart := FALSE;
        prevMixMotorStart := FALSE;
        RETURN;
    END_IF;

    IF NOT opeMode THEN
        State := AUTO_IDLE;

        IF valveAStart AND NOT prevValveAStart THEN
            valveAToggled := NOT valveAToggled;
        END_IF;
        IF valveBStart AND NOT prevValveBStart THEN
            valveBToggled := NOT valveBToggled;
        END_IF;
        IF valveCStart AND NOT prevValveCStart THEN
            valveCToggled := NOT valveCToggled;
        END_IF;
        IF valveDStart AND NOT prevValveDStart THEN
            valveDToggled := NOT valveDToggled;
        END_IF;
        IF mixMotorStart AND NOT prevMixMotorStart THEN
            motorToggled := NOT motorToggled;
        END_IF;

        valveARun := valveAToggled;
        valveBRun := valveBToggled;
        valveCRun := valveCToggled;
        valveDRun := valveDToggled;
        mixMotorRun := motorToggled;
    ELSE
        CASE State OF
            AUTO_IDLE:
                valveAToggled := FALSE;
                valveBToggled := FALSE;
                valveCToggled := FALSE;
                valveDToggled := FALSE;
                motorToggled := FALSE;
                IF autoStart AND NOT prevAutoStart THEN
                    State := AUTO_FILL_A;
                END_IF;

            AUTO_FILL_A:
                valveARun := TRUE;
                IF levelSensor >= 50 THEN
                    valveARun := FALSE;
                    State := AUTO_FILL_B;
                END_IF;

            AUTO_FILL_B:
                valveBRun := TRUE;
                IF levelSensor >= 80 THEN
                    valveBRun := FALSE;
                    IF NOT processMode THEN
                        State := AUTO_MIXING;
                    ELSE
                        State := AUTO_FILL_C;
                    END_IF;
                END_IF;

            AUTO_FILL_C:
                valveCRun := TRUE;
                IF levelSensor >= 100 THEN
                    valveCRun := FALSE;
                    State := AUTO_MIXING;
                END_IF;

            AUTO_MIXING:
                mixMotorRun := TRUE;
                IF mixMotorComplete THEN
                    mixMotorRun := FALSE;
                    State := AUTO_DRAIN;
                END_IF;

            AUTO_DRAIN:
                valveDRun := TRUE;
        END_CASE;
    END_IF;

    prevAutoStart := autoStart;
    prevValveAStart := valveAStart;
    prevValveBStart := valveBStart;
    prevValveCStart := valveCStart;
    prevValveDStart := valveDStart;
    prevMixMotorStart := mixMotorStart;

END_FUNCTION_BLOCK

(* ---- public-hard-02.candidate_01.st ---- *)
FUNCTION_BLOCK FlexibleProcessingControl
VAR_INPUT
    processLength    : USINT;
    sensor1          : BOOL;
    sensor2          : BOOL;
    sensor3          : BOOL;
    sensor4          : BOOL;
    sensor5          : BOOL;
    station1Start    : BOOL;
    station2Complete : BOOL;
    station3Complete : BOOL;
    station4Complete : BOOL;
    processSequence  : ARRAY[1..8] OF USINT;
END_VAR
VAR_OUTPUT
    conveyorLeft  : BOOL;
    conveyorRight : BOOL;
END_VAR
VAR
    state          : (STATE_IDLE, STATE_MOVING);
    currentStep    : USINT;
    targetStation  : USINT;
    currentPosition: USINT;
END_VAR

CASE state OF
STATE_IDLE:
    conveyorLeft  := FALSE;
    conveyorRight := FALSE;
    IF sensor1 AND station1Start AND processLength >= 1 THEN
        currentStep := 1;
        targetStation := processSequence[1];
        state := STATE_MOVING;
    END_IF;

STATE_MOVING:
    IF targetStation > currentPosition THEN
        conveyorRight := TRUE;
        conveyorLeft := FALSE;
        IF sensor2 AND targetStation = 2 THEN
            currentPosition := 2;
        ELSIF sensor3 AND targetStation = 3 THEN
            currentPosition := 3;
        ELSIF sensor4 AND targetStation = 4 THEN
            currentPosition := 4;
        ELSIF sensor5 AND targetStation = 5 THEN
            currentPosition := 5;
        END_IF;
    ELSIF targetStation < currentPosition THEN
        conveyorLeft  := TRUE;
        conveyorRight := FALSE;
        IF sensor4 AND targetStation = 4 THEN
            currentPosition := 4;
        ELSIF sensor3 AND targetStation = 3 THEN
            currentPosition := 3;
        ELSIF sensor2 AND targetStation = 2 THEN
            currentPosition := 2;
        ELSIF sensor1 AND targetStation = 1 THEN
            currentPosition := 1;
        END_IF;
    END_IF;
    IF currentPosition = targetStation THEN
        conveyorLeft  := FALSE;
        conveyorRight := FALSE;
        IF targetStation = 5 THEN
            state := STATE_IDLE;
        ELSE
            IF station2Complete AND targetStation = 2 THEN
                currentStep := currentStep + 1;
                IF currentStep <= processLength THEN
                    targetStation := processSequence[currentStep];
                    state := STATE_MOVING;
                ELSE
                    state := STATE_IDLE;
                END_IF;
            ELSIF station3Complete AND targetStation = 3 THEN
                currentStep := currentStep + 1;
                IF currentStep <= processLength THEN
                    targetStation := processSequence[currentStep];
                    state := STATE_MOVING;
                ELSE
                    state := STATE_IDLE;
                END_IF;
            ELSIF station4Complete AND targetStation = 4 THEN
                currentStep := currentStep + 1;
                IF currentStep <= processLength THEN
                    targetStation := processSequence[currentStep];
                    state := STATE_MOVING;
                ELSE
                    state := STATE_IDLE;
                END_IF;
            END_IF;
        END_IF;
    END_IF;
END_CASE;
END_FUNCTION_BLOCK

(* ---- public-hard-02.raw_candidate_01.st ---- *)
FUNCTION_BLOCK FlexibleProcessingControl
VAR_INPUT
    processLength    : USINT;
    sensor1          : BOOL;
    sensor2          : BOOL;
    sensor3          : BOOL;
    sensor4          : BOOL;
    sensor5          : BOOL;
    station1Start    : BOOL;
    station2Complete : BOOL;
    station3Complete : BOOL;
    station4Complete : BOOL;
    processSequence  : ARRAY[1..8] OF USINT;
END_VAR
VAR_OUTPUT
    conveyorLeft  : BOOL;
    conveyorRight : BOOL;
END_VAR
VAR
    state          : (STATE_IDLE, STATE_MOVING);
    currentStep    : USINT;
    targetStation  : USINT;
    currentPosition: USINT;
END_VAR

CASE state OF
STATE_IDLE:
    conveyorLeft  := FALSE;
    conveyorRight := FALSE;
    IF sensor1 AND station1Start AND processLength >= 1 THEN
        currentStep := 1;
        targetStation := processSequence[1];
        state := STATE_MOVING;
    END_IF

STATE_MOVING:
    IF targetStation > currentPosition THEN
        conveyorRight := TRUE;
        conveyorLeft := FALSE;
        IF sensor2 AND targetStation = 2 THEN
            currentPosition := 2;
        ELSIF sensor3 AND targetStation = 3 THEN
            currentPosition := 3;
        ELSIF sensor4 AND targetStation = 4 THEN
            currentPosition := 4;
        ELSIF sensor5 AND targetStation = 5 THEN
            currentPosition := 5;
        END_IF
    ELSIF targetStation < currentPosition THEN
        conveyorLeft  := TRUE;
        conveyorRight := FALSE;
        IF sensor4 AND targetStation = 4 THEN
            currentPosition := 4;
        ELSIF sensor3 AND targetStation = 3 THEN
            currentPosition := 3;
        ELSIF sensor2 AND targetStation = 2 THEN
            currentPosition := 2;
        ELSIF sensor1 AND targetStation = 1 THEN
            currentPosition := 1;
        END_IF
    END_IF
    IF currentPosition = targetStation THEN
        conveyorLeft  := FALSE;
        conveyorRight := FALSE;
        IF targetStation = 5 THEN
            state := STATE_IDLE;
        ELSE
            IF station2Complete AND targetStation = 2 THEN
                currentStep := currentStep + 1;
                IF currentStep <= processLength THEN
                    targetStation := processSequence[currentStep];
                    state := STATE_MOVING;
                ELSE
                    state := STATE_IDLE;
                END_IF;
            ELSIF station3Complete AND targetStation = 3 THEN
                currentStep := currentStep + 1;
                IF currentStep <= processLength THEN
                    targetStation := processSequence[currentStep];
                    state := STATE_MOVING;
                ELSE
                    state := STATE_IDLE;
                END_IF;
            ELSIF station4Complete AND targetStation = 4 THEN
                currentStep := currentStep + 1;
                IF currentStep <= processLength THEN
                    targetStation := processSequence[currentStep];
                    state := STATE_MOVING;
                ELSE
                    state := STATE_IDLE;
                END_IF;
            END_IF;
        END_IF;
    END_IF;
END_CASE;
END_FUNCTION_BLOCK

(* ---- public-hard-03.candidate_01.st ---- *)
TYPE ST_Recipe :
STRUCT
    recipeID : INT;
    ingredientType : INT;
    ingredientRatio : REAL;
    productionTemperature : REAL;
END_STRUCT;
END_TYPE;

FUNCTION_BLOCK RecipeManagement
VAR_INPUT
    addRecipe : BOOL;
    deleteRecipe : BOOL;
    modifyRecipe : BOOL;
    queryRecipe : BOOL;
    recipeIn : ST_Recipe;
END_VAR
VAR_OUTPUT
    recipeAdded : BOOL := FALSE;
    recipeDeleted : BOOL := FALSE;
    recipeModified : BOOL := FALSE;
    recipeQueryResult : ST_Recipe;
    error : BOOL := FALSE;
    status : WORD := 16#0000;
END_VAR
VAR_IN_OUT
    recipe : ARRAY[1..10] OF ST_Recipe;
END_VAR
VAR
    i : INT;
    foundIndex : INT;
    duplicateExists : BOOL;
    emptySlotIndex : INT;
END_VAR

recipeAdded := FALSE;
recipeDeleted := FALSE;
recipeModified := FALSE;
recipeQueryResult.recipeID := 0;
recipeQueryResult.ingredientType := 0;
recipeQueryResult.ingredientRatio := 0.0;
recipeQueryResult.productionTemperature := 0.0;
error := FALSE;
status := 16#0000;
foundIndex := 0;
duplicateExists := FALSE;
emptySlotIndex := 0;

IF addRecipe THEN
    duplicateExists := FALSE;
    emptySlotIndex := 0;
    FOR i := 1 TO 10 DO
        IF recipe[i].recipeID = recipeIn.recipeID AND recipeIn.recipeID <> 0 THEN
            duplicateExists := TRUE;
            EXIT;
        END_IF;
        IF recipe[i].recipeID = 0 AND emptySlotIndex = 0 THEN
            emptySlotIndex := i;
        END_IF;
    END_FOR;

    IF duplicateExists THEN
        error := TRUE;
        status := 16#8002;
    ELSIF emptySlotIndex = 0 THEN
        error := TRUE;
        status := 16#8003;
    ELSE
        recipe[emptySlotIndex].recipeID := recipeIn.recipeID;
        recipe[emptySlotIndex].ingredientType := recipeIn.ingredientType;
        recipe[emptySlotIndex].ingredientRatio := recipeIn.ingredientRatio;
        recipe[emptySlotIndex].productionTemperature := recipeIn.productionTemperature;
        recipeAdded := TRUE;
    END_IF;
END_IF;

IF deleteRecipe THEN
    foundIndex := 0;
    FOR i := 1 TO 10 DO
        IF recipe[i].recipeID = recipeIn.recipeID THEN
            foundIndex := i;
            EXIT;
        END_IF;
    END_FOR;

    IF foundIndex = 0 THEN
        error := TRUE;
        status := 16#8004;
    ELSE
        recipe[foundIndex].recipeID := 0;
        recipeDeleted := TRUE;
    END_IF;
END_IF;

IF modifyRecipe THEN
    foundIndex := 0;
    FOR i := 1 TO 10 DO
        IF recipe[i].recipeID = recipeIn.recipeID THEN
            foundIndex := i;
            EXIT;
        END_IF;
    END_FOR;

    IF foundIndex = 0 THEN
        error := TRUE;
        status := 16#8005;
    ELSE
        recipe[foundIndex].recipeID := recipeIn.recipeID;
        recipe[foundIndex].ingredientType := recipeIn.ingredientType;
        recipe[foundIndex].ingredientRatio := recipeIn.ingredientRatio;
        recipe[foundIndex].productionTemperature := recipeIn.productionTemperature;
        recipeModified := TRUE;
    END_IF;
END_IF;

IF queryRecipe THEN
    foundIndex := 0;
    FOR i := 1 TO 10 DO
        IF recipe[i].recipeID = recipeIn.recipeID THEN
            foundIndex := i;
            EXIT;
        END_IF;
    END_FOR;

    IF foundIndex = 0 THEN
        error := TRUE;
        status := 16#8001;
    ELSE
        recipeQueryResult.recipeID := recipe[foundIndex].recipeID;
        recipeQueryResult.ingredientType := recipe[foundIndex].ingredientType;
        recipeQueryResult.ingredientRatio := recipe[foundIndex].ingredientRatio;
        recipeQueryResult.productionTemperature := recipe[foundIndex].productionTemperature;
    END_IF;
END_IF;
END_FUNCTION_BLOCK

(* ---- public-hard-03.candidate_02.st ---- *)
TYPE ST_Recipe :
STRUCT
    recipeID : INT;
    ingredientType : INT;
    ingredientRatio : REAL;
    productionTemperature : REAL;
END_STRUCT;
END_TYPE;

FUNCTION_BLOCK RecipeManagement
VAR_INPUT
    addRecipe : BOOL;
    deleteRecipe : BOOL;
    modifyRecipe : BOOL;
    queryRecipe : BOOL;
    recipeIn : ST_Recipe;
END_VAR
VAR_OUTPUT
    recipeAdded : BOOL := FALSE;
    recipeDeleted : BOOL := FALSE;
    recipeModified : BOOL := FALSE;
    recipeQueryResult : ST_Recipe;
    error : BOOL := FALSE;
    status : WORD := 16#0000;
END_VAR
VAR_IN_OUT
    recipe : ARRAY[1..10] OF ST_Recipe;
END_VAR
VAR
    i : INT;
    foundIndex : INT;
    duplicateExists : BOOL;
    emptySlotIndex : INT;
END_VAR

recipeAdded := FALSE;
recipeDeleted := FALSE;
recipeModified := FALSE;
recipeQueryResult.recipeID := 0;
recipeQueryResult.ingredientType := 0;
recipeQueryResult.ingredientRatio := 0.0;
recipeQueryResult.productionTemperature := 0.0;
error := FALSE;
status := 16#0000;
foundIndex := 0;
duplicateExists := FALSE;
emptySlotIndex := 0;

IF addRecipe THEN
    duplicateExists := FALSE;
    emptySlotIndex := 0;
    FOR i := 1 TO 10 DO
        IF recipe[i].recipeID = recipeIn.recipeID AND recipeIn.recipeID <> 0 THEN
            duplicateExists := TRUE;
            EXIT;
        END_IF;
        IF recipe[i].recipeID = 0 AND emptySlotIndex = 0 THEN
            emptySlotIndex := i;
        END_IF;
    END_FOR;

    IF duplicateExists THEN
        error := TRUE;
        status := 16#8002;
    ELSIF emptySlotIndex = 0 THEN
        error := TRUE;
        status := 16#8003;
    ELSE
        recipe[emptySlotIndex].recipeID := recipeIn.recipeID;
        recipe[emptySlotIndex].ingredientType := recipeIn.ingredientType;
        recipe[emptySlotIndex].ingredientRatio := recipeIn.ingredientRatio;
        recipe[emptySlotIndex].productionTemperature := recipeIn.productionTemperature;
        recipeAdded := TRUE;
    END_IF;
END_IF;

IF deleteRecipe THEN
    foundIndex := 0;
    FOR i := 1 TO 10 DO
        IF recipe[i].recipeID = recipeIn.recipeID THEN
            foundIndex := i;
            EXIT;
        END_IF;
    END_FOR;

    IF foundIndex = 0 THEN
        error := TRUE;
        status := 16#8004;
    ELSE
        recipe[foundIndex].recipeID := 0;
        recipeDeleted := TRUE;
    END_IF;
END_IF;

IF modifyRecipe THEN
    foundIndex := 0;
    FOR i := 1 TO 10 DO
        IF recipe[i].recipeID = recipeIn.recipeID THEN
            foundIndex := i;
            EXIT;
        END_IF;
    END_FOR;

    IF foundIndex = 0 THEN
        error := TRUE;
        status := 16#8005;
    ELSE
        recipe[foundIndex].recipeID := recipeIn.recipeID;
        recipe[foundIndex].ingredientType := recipeIn.ingredientType;
        recipe[foundIndex].ingredientRatio := recipeIn.ingredientRatio;
        recipe[foundIndex].productionTemperature := recipeIn.productionTemperature;
        recipeModified := TRUE;
    END_IF;
END_IF;

IF queryRecipe THEN
    foundIndex := 0;
    FOR i := 1 TO 10 DO
        IF recipe[i].recipeID = recipeIn.recipeID THEN
            foundIndex := i;
            EXIT;
        END_IF;
    END_FOR;

    IF foundIndex = 0 THEN
        error := TRUE;
        status := 16#8001;
    ELSE
        recipeQueryResult.recipeID := recipe[foundIndex].recipeID;
        recipeQueryResult.ingredientType := recipe[foundIndex].ingredientType;
        recipeQueryResult.ingredientRatio := recipe[foundIndex].ingredientRatio;
        recipeQueryResult.productionTemperature := recipe[foundIndex].productionTemperature;
    END_IF;
END_IF;
END_FUNCTION_BLOCK

(* ---- public-hard-03.raw_candidate_01.st ---- *)
TYPE ST_Recipe :
STRUCT
    recipeID : INT;
    ingredientType : INT;
    ingredientRatio : REAL;
    productionTemperature : REAL;
END_STRUCT
END_TYPE

FUNCTION_BLOCK RecipeManagement
VAR_INPUT
    addRecipe : BOOL;
    deleteRecipe : BOOL;
    modifyRecipe : BOOL;
    queryRecipe : BOOL;
    recipeIn : ST_Recipe;
END_VAR
VAR_OUTPUT
    recipeAdded : BOOL := FALSE;
    recipeDeleted : BOOL := FALSE;
    recipeModified : BOOL := FALSE;
    recipeQueryResult : ST_Recipe;
    error : BOOL := FALSE;
    status : WORD := 16#0000;
END_VAR
VAR_IN_OUT
    recipe : ARRAY[1..10] OF ST_Recipe;
END_VAR
VAR
    i : INT;
    foundIndex : INT;
    duplicateExists : BOOL;
    emptySlotIndex : INT;
END_VAR

recipeAdded := FALSE;
recipeDeleted := FALSE;
recipeModified := FALSE;
recipeQueryResult.recipeID := 0;
recipeQueryResult.ingredientType := 0;
recipeQueryResult.ingredientRatio := 0.0;
recipeQueryResult.productionTemperature := 0.0;
error := FALSE;
status := 16#0000;
foundIndex := 0;
duplicateExists := FALSE;
emptySlotIndex := 0;

IF addRecipe THEN
    duplicateExists := FALSE;
    emptySlotIndex := 0;
    FOR i := 1 TO 10 DO
        IF recipe[i].recipeID = recipeIn.recipeID AND recipeIn.recipeID <> 0 THEN
            duplicateExists := TRUE;
            EXIT;
        END_IF
        IF recipe[i].recipeID = 0 AND emptySlotIndex = 0 THEN
            emptySlotIndex := i;
        END_IF
    END_FOR;

    IF duplicateExists THEN
        error := TRUE;
        status := 16#8002;
    ELSIF emptySlotIndex = 0 THEN
        error := TRUE;
        status := 16#8003;
    ELSE
        recipe[emptySlotIndex].recipeID := recipeIn.recipeID;
        recipe[emptySlotIndex].ingredientType := recipeIn.ingredientType;
        recipe[emptySlotIndex].ingredientRatio := recipeIn.ingredientRatio;
        recipe[emptySlotIndex].productionTemperature := recipeIn.productionTemperature;
        recipeAdded := TRUE;
    END_IF;
END_IF;

IF deleteRecipe THEN
    foundIndex := 0;
    FOR i := 1 TO 10 DO
        IF recipe[i].recipeID = recipeIn.recipeID THEN
            foundIndex := i;
            EXIT;
        END_IF
    END_FOR;

    IF foundIndex = 0 THEN
        error := TRUE;
        status := 16#8004;
    ELSE
        recipe[foundIndex].recipeID := 0;
        recipeDeleted := TRUE;
    END_IF;
END_IF;

IF modifyRecipe THEN
    foundIndex := 0;
    FOR i := 1 TO 10 DO
        IF recipe[i].recipeID = recipeIn.recipeID THEN
            foundIndex := i;
            EXIT;
        END_IF
    END_FOR;

    IF foundIndex = 0 THEN
        error := TRUE;
        status := 16#8005;
    ELSE
        recipe[foundIndex].recipeID := recipeIn.recipeID;
        recipe[foundIndex].ingredientType := recipeIn.ingredientType;
        recipe[foundIndex].ingredientRatio := recipeIn.ingredientRatio;
        recipe[foundIndex].productionTemperature := recipeIn.productionTemperature;
        recipeModified := TRUE;
    END_IF;
END_IF;

IF queryRecipe THEN
    foundIndex := 0;
    FOR i := 1 TO 10 DO
        IF recipe[i].recipeID = recipeIn.recipeID THEN
            foundIndex := i;
            EXIT;
        END_IF
    END_FOR;

    IF foundIndex = 0 THEN
        error := TRUE;
        status := 16#8001;
    ELSE
        recipeQueryResult.recipeID := recipe[foundIndex].recipeID;
        recipeQueryResult.ingredientType := recipe[foundIndex].ingredientType;
        recipeQueryResult.ingredientRatio := recipe[foundIndex].ingredientRatio;
        recipeQueryResult.productionTemperature := recipe[foundIndex].productionTemperature;
    END_IF;
END_IF;
END_FUNCTION_BLOCK

(* ---- public-hard-03.raw_candidate_02.st ---- *)
TYPE ST_Recipe :
STRUCT
    recipeID : INT;
    ingredientType : INT;
    ingredientRatio : REAL;
    productionTemperature : REAL;
END_STRUCT
END_TYPE

FUNCTION_BLOCK RecipeManagement
VAR_INPUT
    addRecipe : BOOL;
    deleteRecipe : BOOL;
    modifyRecipe : BOOL;
    queryRecipe : BOOL;
    recipeIn : ST_Recipe;
END_VAR
VAR_OUTPUT
    recipeAdded : BOOL := FALSE;
    recipeDeleted : BOOL := FALSE;
    recipeModified : BOOL := FALSE;
    recipeQueryResult : ST_Recipe;
    error : BOOL := FALSE;
    status : WORD := 16#0000;
END_VAR
VAR_IN_OUT
    recipe : ARRAY[1..10] OF ST_Recipe;
END_VAR
VAR
    i : INT;
    foundIndex : INT;
    duplicateExists : BOOL;
    emptySlotIndex : INT;
END_VAR

recipeAdded := FALSE;
recipeDeleted := FALSE;
recipeModified := FALSE;
recipeQueryResult.recipeID := 0;
recipeQueryResult.ingredientType := 0;
recipeQueryResult.ingredientRatio := 0.0;
recipeQueryResult.productionTemperature := 0.0;
error := FALSE;
status := 16#0000;
foundIndex := 0;
duplicateExists := FALSE;
emptySlotIndex := 0;

IF addRecipe THEN
    duplicateExists := FALSE;
    emptySlotIndex := 0;
    FOR i := 1 TO 10 DO
        IF recipe[i].recipeID = recipeIn.recipeID AND recipeIn.recipeID <> 0 THEN
            duplicateExists := TRUE;
            EXIT;
        END_IF;
        IF recipe[i].recipeID = 0 AND emptySlotIndex = 0 THEN
            emptySlotIndex := i;
        END_IF;
    END_FOR;

    IF duplicateExists THEN
        error := TRUE;
        status := 16#8002;
    ELSIF emptySlotIndex = 0 THEN
        error := TRUE;
        status := 16#8003;
    ELSE
        recipe[emptySlotIndex].recipeID := recipeIn.recipeID;
        recipe[emptySlotIndex].ingredientType := recipeIn.ingredientType;
        recipe[emptySlotIndex].ingredientRatio := recipeIn.ingredientRatio;
        recipe[emptySlotIndex].productionTemperature := recipeIn.productionTemperature;
        recipeAdded := TRUE;
    END_IF;
END_IF;

IF deleteRecipe THEN
    foundIndex := 0;
    FOR i := 1 TO 10 DO
        IF recipe[i].recipeID = recipeIn.recipeID THEN
            foundIndex := i;
            EXIT;
        END_IF;
    END_FOR;

    IF foundIndex = 0 THEN
        error := TRUE;
        status := 16#8004;
    ELSE
        recipe[foundIndex].recipeID := 0;
        recipeDeleted := TRUE;
    END_IF;
END_IF;

IF modifyRecipe THEN
    foundIndex := 0;
    FOR i := 1 TO 10 DO
        IF recipe[i].recipeID = recipeIn.recipeID THEN
            foundIndex := i;
            EXIT;
        END_IF;
    END_FOR;

    IF foundIndex = 0 THEN
        error := TRUE;
        status := 16#8005;
    ELSE
        recipe[foundIndex].recipeID := recipeIn.recipeID;
        recipe[foundIndex].ingredientType := recipeIn.ingredientType;
        recipe[foundIndex].ingredientRatio := recipeIn.ingredientRatio;
        recipe[foundIndex].productionTemperature := recipeIn.productionTemperature;
        recipeModified := TRUE;
    END_IF;
END_IF;

IF queryRecipe THEN
    foundIndex := 0;
    FOR i := 1 TO 10 DO
        IF recipe[i].recipeID = recipeIn.recipeID THEN
            foundIndex := i;
            EXIT;
        END_IF;
    END_FOR;

    IF foundIndex = 0 THEN
        error := TRUE;
        status := 16#8001;
    ELSE
        recipeQueryResult.recipeID := recipe[foundIndex].recipeID;
        recipeQueryResult.ingredientType := recipe[foundIndex].ingredientType;
        recipeQueryResult.ingredientRatio := recipe[foundIndex].ingredientRatio;
        recipeQueryResult.productionTemperature := recipe[foundIndex].productionTemperature;
    END_IF;
END_IF;
END_FUNCTION_BLOCK

(* ---- public-hard-04.candidate_01.st ---- *)
FUNCTION_BLOCK FB_FIFO_Queue
VAR_INPUT
    enqueue  : BOOL;
    dequeue  : BOOL;
    reset    : BOOL;
END_VAR
VAR_OUTPUT
    elementCount : DINT := 0;
    status       : WORD := 16#0000;
END_VAR
VAR_IN_OUT
    item   : VARIANT;
    buffer : VARIANT;
END_VAR
VAR
    head         : DINT := 0;
    tail         : DINT := 0;
    capacity     : DINT := 0;
    prevEnqueue  : BOOL := FALSE;
    prevDequeue  : BOOL := FALSE;
    initDone     : BOOL := FALSE;
END_VAR

// Initialize capacity from buffer array bounds on first invocation
IF NOT initDone THEN
    capacity := __GETUPPERBOUND(buffer, 1) + 1;
    initDone := TRUE;
END_IF;

// Reset takes priority over all other operations
IF reset THEN
    head := 0;
    tail := 0;
    elementCount := 0;
    status := 16#0000;
    prevEnqueue := FALSE;
    prevDequeue := FALSE;
    RETURN;
END_IF;

// Rising edge detection for enqueue
IF enqueue AND NOT prevEnqueue THEN
    prevEnqueue := TRUE;
    IF elementCount >= capacity THEN
        status := 16#8002;
    ELSE
        __SETATINDEX(buffer, tail, item);
        tail := (tail + 1) MOD capacity;
        elementCount := elementCount + 1;
        status := 16#0000;
    END_IF;
ELSE
    prevEnqueue := enqueue;
END_IF;

// Rising edge detection for dequeue
IF dequeue AND NOT prevDequeue THEN
    prevDequeue := TRUE;
    IF elementCount <= 0 THEN
        status := 16#8001;
    ELSE
        item := __GETATINDEX(buffer, head);
        head := (head + 1) MOD capacity;
        elementCount := elementCount - 1;
        status := 16#0000;
    END_IF;
ELSE
    prevDequeue := dequeue;
END_IF;

// Set status to no-error if no operation was performed this cycle
IF NOT reset AND NOT (enqueue AND NOT prevEnqueue) AND NOT (dequeue AND NOT prevDequeue) THEN
    status := 16#0000;
END_IF;

END_FUNCTION_BLOCK

(* ---- public-hard-04.candidate_02.st ---- *)
FUNCTION_BLOCK FB_FIFO_Queue
VAR_INPUT
    enqueue  : BOOL;
    dequeue  : BOOL;
    reset    : BOOL;
END_VAR
VAR_OUTPUT
    elementCount : DINT := 0;
    status       : WORD := 16#0000;
END_VAR
VAR_IN_OUT
    item   : VARIANT;
    buffer : VARIANT;
END_VAR
VAR
    head         : DINT := 0;
    tail         : DINT := 0;
    capacity     : DINT := 0;
    prevEnqueue  : BOOL := FALSE;
    prevDequeue  : BOOL := FALSE;
    initDone     : BOOL := FALSE;
END_VAR

// Initialize capacity from buffer array bounds on first invocation
IF NOT initDone THEN
    capacity := __GETUPPERBOUND(buffer, 1) + 1;
    initDone := TRUE;
END_IF;

// Reset takes priority over all other operations
IF reset THEN
    head := 0;
    tail := 0;
    elementCount := 0;
    status := 16#0000;
    prevEnqueue := FALSE;
    prevDequeue := FALSE;
    RETURN;
END_IF;

// Rising edge detection for enqueue
IF enqueue AND NOT prevEnqueue THEN
    prevEnqueue := TRUE;
    IF elementCount >= capacity THEN
        status := 16#8002;
    ELSE
        __SETATINDEX(buffer, tail, item);
        tail := (tail + 1) MOD capacity;
        elementCount := elementCount + 1;
        status := 16#0000;
    END_IF;
ELSE
    prevEnqueue := enqueue;
END_IF;

// Rising edge detection for dequeue
IF dequeue AND NOT prevDequeue THEN
    prevDequeue := TRUE;
    IF elementCount <= 0 THEN
        status := 16#8001;
    ELSE
        item := __GETATINDEX(buffer, head);
        head := (head + 1) MOD capacity;
        elementCount := elementCount - 1;
        status := 16#0000;
    END_IF;
ELSE
    prevDequeue := dequeue;
END_IF;

// Set status to no-error if no operation was performed this cycle
IF NOT reset AND NOT (enqueue AND NOT prevEnqueue) AND NOT (dequeue AND NOT prevDequeue) THEN
    status := 16#0000;
END_IF;

END_FUNCTION_BLOCK

(* ---- public-hard-04.raw_candidate_01.st ---- *)
FUNCTION_BLOCK FB_FIFO_Queue
VAR_INPUT
    enqueue  : BOOL;
    dequeue  : BOOL;
    reset    : BOOL;
END_VAR
VAR_OUTPUT
    elementCount : DINT := 0;
    status       : WORD := 16#0000;
END_VAR
VAR_IN_OUT
    item   : VARIANT;
    buffer : VARIANT;
END_VAR
VAR
    head         : DINT := 0;
    tail         : DINT := 0;
    capacity     : DINT := 0;
    prevEnqueue  : BOOL := FALSE;
    prevDequeue  : BOOL := FALSE;
    initDone     : BOOL := FALSE;
END_VAR

// Initialize capacity from buffer array bounds on first invocation
IF NOT initDone THEN
    capacity := __GETUPPERBOUND(buffer, 1) + 1;
    initDone := TRUE;
END_IF

// Reset takes priority over all other operations
IF reset THEN
    head := 0;
    tail := 0;
    elementCount := 0;
    status := 16#0000;
    prevEnqueue := FALSE;
    prevDequeue := FALSE;
    RETURN;
END_IF;

// Rising edge detection for enqueue
IF enqueue AND NOT prevEnqueue THEN
    prevEnqueue := TRUE;
    IF elementCount >= capacity THEN
        status := 16#8002;
    ELSE
        __SETATINDEX(buffer, tail, item);
        tail := (tail + 1) MOD capacity;
        elementCount := elementCount + 1;
        status := 16#0000;
    END_IF;
ELSE
    prevEnqueue := enqueue;
END_IF;

// Rising edge detection for dequeue
IF dequeue AND NOT prevDequeue THEN
    prevDequeue := TRUE;
    IF elementCount <= 0 THEN
        status := 16#8001;
    ELSE
        item := __GETATINDEX(buffer, head);
        head := (head + 1) MOD capacity;
        elementCount := elementCount - 1;
        status := 16#0000;
    END_IF;
ELSE
    prevDequeue := dequeue;
END_IF;

// Set status to no-error if no operation was performed this cycle
IF NOT reset AND NOT (enqueue AND NOT prevEnqueue) AND NOT (dequeue AND NOT prevDequeue) THEN
    status := 16#0000;
END_IF;

END_FUNCTION_BLOCK

(* ---- public-hard-04.raw_candidate_02.st ---- *)
FUNCTION_BLOCK FB_FIFO_Queue
VAR_INPUT
    enqueue  : BOOL;
    dequeue  : BOOL;
    reset    : BOOL;
END_VAR
VAR_OUTPUT
    elementCount : DINT := 0;
    status       : WORD := 16#0000;
END_VAR
VAR_IN_OUT
    item   : VARIANT;
    buffer : VARIANT;
END_VAR
VAR
    head         : DINT := 0;
    tail         : DINT := 0;
    capacity     : DINT := 0;
    prevEnqueue  : BOOL := FALSE;
    prevDequeue  : BOOL := FALSE;
    initDone     : BOOL := FALSE;
END_VAR

// Initialize capacity from buffer array bounds on first invocation
IF NOT initDone THEN
    capacity := __GETUPPERBOUND(buffer, 1) + 1;
    initDone := TRUE;
END_IF;

// Reset takes priority over all other operations
IF reset THEN
    head := 0;
    tail := 0;
    elementCount := 0;
    status := 16#0000;
    prevEnqueue := FALSE;
    prevDequeue := FALSE;
    RETURN;
END_IF;

// Rising edge detection for enqueue
IF enqueue AND NOT prevEnqueue THEN
    prevEnqueue := TRUE;
    IF elementCount >= capacity THEN
        status := 16#8002;
    ELSE
        __SETATINDEX(buffer, tail, item);
        tail := (tail + 1) MOD capacity;
        elementCount := elementCount + 1;
        status := 16#0000;
    END_IF;
ELSE
    prevEnqueue := enqueue;
END_IF;

// Rising edge detection for dequeue
IF dequeue AND NOT prevDequeue THEN
    prevDequeue := TRUE;
    IF elementCount <= 0 THEN
        status := 16#8001;
    ELSE
        item := __GETATINDEX(buffer, head);
        head := (head + 1) MOD capacity;
        elementCount := elementCount - 1;
        status := 16#0000;
    END_IF;
ELSE
    prevDequeue := dequeue;
END_IF;

// Set status to no-error if no operation was performed this cycle
IF NOT reset AND NOT (enqueue AND NOT prevEnqueue) AND NOT (dequeue AND NOT prevDequeue) THEN
    status := 16#0000;
END_IF;

END_FUNCTION_BLOCK

(* ---- public-hard-05.candidate_01.st ---- *)
FUNCTION_BLOCK MechanicalArmControl
VAR_INPUT
    ManualMode       : BOOL;
    SingleStepMode   : BOOL;
    SingleCycleMode  : BOOL;
    ContinuousMode   : BOOL;
    EmergencyStop    : BOOL;
    Start            : BOOL;
    DownButton       : BOOL;
    UpButton         : BOOL;
    LeftButton       : BOOL;
    RightButton      : BOOL;
    GripButton       : BOOL;
    ReleaseButton    : BOOL;
    DownLimitSwitch  : BOOL;
    UpLimitSwitch    : BOOL;
    LeftLimitSwitch  : BOOL;
    RightLimitSwitch : BOOL;
    GripLimitSwitch  : BOOL;
    ReleaseLimitSwitch : BOOL;
END_VAR

VAR_OUTPUT
    MoveDown       : BOOL;
    MoveUp         : BOOL;
    MoveLeft       : BOOL;
    MoveRight      : BOOL;
    ActivateGrip   : BOOL;
    ActivateRelease : BOOL;
END_VAR

VAR
    step        : UINT;
    prevStart   : BOOL;
    startPressed : BOOL;
    prevStep    : UINT;
    cycleActive : BOOL;
END_VAR

// Emergency stop handling
IF NOT EmergencyStop THEN
    MoveDown := FALSE;
    MoveUp := FALSE;
    MoveLeft := FALSE;
    MoveRight := FALSE;
    ActivateGrip := FALSE;
    ActivateRelease := FALSE;
    step := 0;
    prevStep := 0;
    cycleActive := FALSE;
    RETURN;
END_IF;

// Detect rising edge of Start
startPressed := Start AND NOT prevStart;
prevStart := Start;

// Manual mode: Direct button control, stop at limit switches
IF ManualMode THEN
    MoveDown := DownButton AND NOT DownLimitSwitch;
    MoveUp := UpButton AND NOT UpLimitSwitch;
    MoveLeft := LeftButton AND NOT LeftLimitSwitch;
    MoveRight := RightButton AND NOT RightLimitSwitch;
    ActivateGrip := GripButton;
    ActivateRelease := ReleaseButton;
    step := 0;
    cycleActive := FALSE;

// Single step mode: One action per Start press, wait for completion
ELSIF SingleStepMode THEN
    IF startPressed THEN
        step := step + 1;
        IF step > 8 THEN
            step := 1;
        END_IF;
        prevStep := step;
    END_IF;

    CASE step OF
        1: MoveDown := NOT DownLimitSwitch;
        2: ActivateGrip := NOT GripLimitSwitch;
        3: MoveUp := NOT UpLimitSwitch;
        4: MoveRight := NOT RightLimitSwitch;
        5: MoveDown := NOT DownLimitSwitch;
        6: ActivateRelease := NOT ReleaseLimitSwitch;
        7: MoveUp := NOT UpLimitSwitch;
        8: MoveLeft := NOT LeftLimitSwitch;
    END_CASE;

    IF step <> prevStep THEN
        prevStep := step;
    ELSIF step > 0 THEN
        CASE step OF
            1: IF DownLimitSwitch THEN step := 0; prevStep := 0; END_IF;
            2: IF GripLimitSwitch THEN step := 0; prevStep := 0; END_IF;
            3: IF UpLimitSwitch THEN step := 0; prevStep := 0; END_IF;
            4: IF RightLimitSwitch THEN step := 0; prevStep := 0; END_IF;
            5: IF DownLimitSwitch THEN step := 0; prevStep := 0; END_IF;
            6: IF ReleaseLimitSwitch THEN step := 0; prevStep := 0; END_IF;
            7: IF UpLimitSwitch THEN step := 0; prevStep := 0; END_IF;
            8: IF LeftLimitSwitch THEN step := 0; prevStep := 0; END_IF;
        END_CASE;
    END_IF;

// Single cycle mode: Full sequence automatic, stop at end
ELSIF SingleCycleMode THEN
    IF startPressed THEN
        cycleActive := TRUE;
        prevStep := 0;
    END_IF;

    IF cycleActive THEN
        CASE step OF
            0: MoveDown := NOT DownLimitSwitch;
            1: ActivateGrip := NOT GripLimitSwitch;
            2: MoveUp := NOT UpLimitSwitch;
            3: MoveRight := NOT RightLimitSwitch;
            4: MoveDown := NOT DownLimitSwitch;
            5: ActivateRelease := NOT ReleaseLimitSwitch;
            6: MoveUp := NOT UpLimitSwitch;
            7: MoveLeft := NOT LeftLimitSwitch;
        END_CASE;

        IF step <> prevStep THEN
            prevStep := step;
        ELSIF step < 8 THEN
            CASE step OF
                0: IF DownLimitSwitch THEN step := 1; prevStep := 1; END_IF;
                1: IF GripLimitSwitch THEN step := 2; prevStep := 2; END_IF;
                2: IF UpLimitSwitch THEN step := 3; prevStep := 3; END_IF;
                3: IF RightLimitSwitch THEN step := 4; prevStep := 4; END_IF;
                4: IF DownLimitSwitch THEN step := 5; prevStep := 5; END_IF;
                5: IF ReleaseLimitSwitch THEN step := 6; prevStep := 6; END_IF;
                6: IF UpLimitSwitch THEN step := 7; prevStep := 7; END_IF;
                7: IF LeftLimitSwitch THEN step := 0; prevStep := 0; cycleActive := FALSE; END_IF;
            END_CASE;
        END_IF;
    END_IF;

// Continuous mode: Full sequence repeating
ELSIF ContinuousMode THEN
    IF startPressed THEN
        cycleActive := TRUE;
        prevStep := 0;
    END_IF;

    IF cycleActive THEN
        CASE step OF
            0: MoveDown := NOT DownLimitSwitch;
            1: ActivateGrip := NOT GripLimitSwitch;
            2: MoveUp := NOT UpLimitSwitch;
            3: MoveRight := NOT RightLimitSwitch;
            4: MoveDown := NOT DownLimitSwitch;
            5: ActivateRelease := NOT ReleaseLimitSwitch;
            6: MoveUp := NOT UpLimitSwitch;
            7: MoveLeft := NOT LeftLimitSwitch;
        END_CASE;

        IF step <> prevStep THEN
            prevStep := step;
        ELSIF step < 8 THEN
            CASE step OF
                0: IF DownLimitSwitch THEN step := 1; prevStep := 1; END_IF;
                1: IF GripLimitSwitch THEN step := 2; prevStep := 2; END_IF;
                2: IF UpLimitSwitch THEN step := 3; prevStep := 3; END_IF;
                3: IF RightLimitSwitch THEN step := 4; prevStep := 4; END_IF;
                4: IF DownLimitSwitch THEN step := 5; prevStep := 5; END_IF;
                5: IF ReleaseLimitSwitch THEN step := 6; prevStep := 6; END_IF;
                6: IF UpLimitSwitch THEN step := 7; prevStep := 7; END_IF;
                7: IF LeftLimitSwitch THEN step := 0; prevStep := 0; END_IF;
            END_CASE;
        END_IF;
    END_IF;

END_IF;
END_FUNCTION_BLOCK

(* ---- public-hard-05.candidate_02.st ---- *)
FUNCTION_BLOCK MechanicalArmControl
VAR_INPUT
    ManualMode       : BOOL;
    SingleStepMode   : BOOL;
    SingleCycleMode  : BOOL;
    ContinuousMode   : BOOL;
    EmergencyStop    : BOOL;
    Start            : BOOL;
    DownButton       : BOOL;
    UpButton         : BOOL;
    LeftButton       : BOOL;
    RightButton      : BOOL;
    GripButton       : BOOL;
    ReleaseButton    : BOOL;
    DownLimitSwitch  : BOOL;
    UpLimitSwitch    : BOOL;
    LeftLimitSwitch  : BOOL;
    RightLimitSwitch : BOOL;
    GripLimitSwitch  : BOOL;
    ReleaseLimitSwitch : BOOL;
END_VAR

VAR_OUTPUT
    MoveDown       : BOOL;
    MoveUp         : BOOL;
    MoveLeft       : BOOL;
    MoveRight      : BOOL;
    ActivateGrip   : BOOL;
    ActivateRelease : BOOL;
END_VAR

VAR
    step         : UINT;
    prevStart    : BOOL;
    startPressed : BOOL;
    cycleActive  : BOOL;
END_VAR

// Reset all outputs first
MoveDown := FALSE;
MoveUp := FALSE;
MoveLeft := FALSE;
MoveRight := FALSE;
ActivateGrip := FALSE;
ActivateRelease := FALSE;

// Emergency stop: immediate halt
IF NOT EmergencyStop THEN
    step := 0;
    cycleActive := FALSE;
    prevStart := FALSE;
    RETURN;
END_IF;

// Rising edge detection for Start
startPressed := Start AND NOT prevStart;
prevStart := Start;

// Manual mode: Direct control via buttons
IF ManualMode THEN
    MoveDown := DownButton AND NOT DownLimitSwitch;
    MoveUp := UpButton AND NOT UpLimitSwitch;
    MoveLeft := LeftButton AND NOT LeftLimitSwitch;
    MoveRight := RightButton AND NOT RightLimitSwitch;
    ActivateGrip := GripButton;
    ActivateRelease := ReleaseButton;
    step := 0;
    cycleActive := FALSE;

// Single step mode: One action per Start press
ELSIF SingleStepMode THEN
    IF startPressed THEN
        step := step + 1;
        IF step > 8 THEN
            step := 1;
        END_IF;
    END_IF;

    // Execute current step
    CASE step OF
        1: MoveDown := NOT DownLimitSwitch;
        2: ActivateGrip := NOT GripLimitSwitch;
        3: MoveUp := NOT UpLimitSwitch;
        4: MoveRight := NOT RightLimitSwitch;
        5: MoveDown := NOT DownLimitSwitch;
        6: ActivateRelease := NOT ReleaseLimitSwitch;
        7: MoveUp := NOT UpLimitSwitch;
        8: MoveLeft := NOT LeftLimitSwitch;
    END_CASE;

    // Check completion and reset to wait for next Start
    CASE step OF
        1: IF DownLimitSwitch THEN step := 0; END_IF;
        2: IF GripLimitSwitch THEN step := 0; END_IF;
        3: IF UpLimitSwitch THEN step := 0; END_IF;
        4: IF RightLimitSwitch THEN step := 0; END_IF;
        5: IF DownLimitSwitch THEN step := 0; END_IF;
        6: IF ReleaseLimitSwitch THEN step := 0; END_IF;
        7: IF UpLimitSwitch THEN step := 0; END_IF;
        8: IF LeftLimitSwitch THEN step := 0; END_IF;
    END_CASE;

// Single cycle mode: Full sequence automatic, stop at end
ELSIF SingleCycleMode THEN
    IF startPressed THEN
        step := 0;
        cycleActive := TRUE;
    END_IF;

    IF cycleActive THEN
        CASE step OF
            0: MoveDown := NOT DownLimitSwitch;
            1: ActivateGrip := NOT GripLimitSwitch;
            2: MoveUp := NOT UpLimitSwitch;
            3: MoveRight := NOT RightLimitSwitch;
            4: MoveDown := NOT DownLimitSwitch;
            5: ActivateRelease := NOT ReleaseLimitSwitch;
            6: MoveUp := NOT UpLimitSwitch;
            7: MoveLeft := NOT LeftLimitSwitch;
        END_CASE;

        CASE step OF
            0: IF DownLimitSwitch THEN step := 1; END_IF;
            1: IF GripLimitSwitch THEN step := 2; END_IF;
            2: IF UpLimitSwitch THEN step := 3; END_IF;
            3: IF RightLimitSwitch THEN step := 4; END_IF;
            4: IF DownLimitSwitch THEN step := 5; END_IF;
            5: IF ReleaseLimitSwitch THEN step := 6; END_IF;
            6: IF UpLimitSwitch THEN step := 7; END_IF;
            7: IF LeftLimitSwitch THEN
                   step := 0;
                   cycleActive := FALSE;
               END_IF;
        END_CASE;
    END_IF;

// Continuous mode: Full sequence repeating
ELSIF ContinuousMode THEN
    IF startPressed THEN
        step := 0;
        cycleActive := TRUE;
    END_IF;

    IF cycleActive THEN
        CASE step OF
            0: MoveDown := NOT DownLimitSwitch;
            1: ActivateGrip := NOT GripLimitSwitch;
            2: MoveUp := NOT UpLimitSwitch;
            3: MoveRight := NOT RightLimitSwitch;
            4: MoveDown := NOT DownLimitSwitch;
            5: ActivateRelease := NOT ReleaseLimitSwitch;
            6: MoveUp := NOT UpLimitSwitch;
            7: MoveLeft := NOT LeftLimitSwitch;
        END_CASE;

        CASE step OF
            0: IF DownLimitSwitch THEN step := 1; END_IF;
            1: IF GripLimitSwitch THEN step := 2; END_IF;
            2: IF UpLimitSwitch THEN step := 3; END_IF;
            3: IF RightLimitSwitch THEN step := 4; END_IF;
            4: IF DownLimitSwitch THEN step := 5; END_IF;
            5: IF ReleaseLimitSwitch THEN step := 6; END_IF;
            6: IF UpLimitSwitch THEN step := 7; END_IF;
            7: IF LeftLimitSwitch THEN step := 0; END_IF;
        END_CASE;
    END_IF;

END_IF;
END_FUNCTION_BLOCK

(* ---- public-hard-05.raw_candidate_01.st ---- *)
FUNCTION_BLOCK MechanicalArmControl
VAR_INPUT
    ManualMode       : BOOL;
    SingleStepMode   : BOOL;
    SingleCycleMode  : BOOL;
    ContinuousMode   : BOOL;
    EmergencyStop    : BOOL;
    Start            : BOOL;
    DownButton       : BOOL;
    UpButton         : BOOL;
    LeftButton       : BOOL;
    RightButton      : BOOL;
    GripButton       : BOOL;
    ReleaseButton    : BOOL;
    DownLimitSwitch  : BOOL;
    UpLimitSwitch    : BOOL;
    LeftLimitSwitch  : BOOL;
    RightLimitSwitch : BOOL;
    GripLimitSwitch  : BOOL;
    ReleaseLimitSwitch : BOOL;
END_VAR

VAR_OUTPUT
    MoveDown       : BOOL;
    MoveUp         : BOOL;
    MoveLeft       : BOOL;
    MoveRight      : BOOL;
    ActivateGrip   : BOOL;
    ActivateRelease : BOOL;
END_VAR

VAR
    step        : UINT;
    prevStart   : BOOL;
    startPressed : BOOL;
    prevStep    : UINT;
    cycleActive : BOOL;
END_VAR

// Emergency stop handling
IF NOT EmergencyStop THEN
    MoveDown := FALSE;
    MoveUp := FALSE;
    MoveLeft := FALSE;
    MoveRight := FALSE;
    ActivateGrip := FALSE;
    ActivateRelease := FALSE;
    step := 0;
    prevStep := 0;
    cycleActive := FALSE;
    RETURN;
END_IF;

// Detect rising edge of Start
startPressed := Start AND NOT prevStart;
prevStart := Start;

// Manual mode: Direct button control, stop at limit switches
IF ManualMode THEN
    MoveDown := DownButton AND NOT DownLimitSwitch;
    MoveUp := UpButton AND NOT UpLimitSwitch;
    MoveLeft := LeftButton AND NOT LeftLimitSwitch;
    MoveRight := RightButton AND NOT RightLimitSwitch;
    ActivateGrip := GripButton;
    ActivateRelease := ReleaseButton;
    step := 0;
    cycleActive := FALSE;

// Single step mode: One action per Start press, wait for completion
ELSIF SingleStepMode THEN
    IF startPressed THEN
        step := step + 1;
        IF step > 8 THEN
            step := 1;
        END_IF;
        prevStep := step;
    END_IF;

    CASE step OF
        1: MoveDown := NOT DownLimitSwitch;
        2: ActivateGrip := NOT GripLimitSwitch;
        3: MoveUp := NOT UpLimitSwitch;
        4: MoveRight := NOT RightLimitSwitch;
        5: MoveDown := NOT DownLimitSwitch;
        6: ActivateRelease := NOT ReleaseLimitSwitch;
        7: MoveUp := NOT UpLimitSwitch;
        8: MoveLeft := NOT LeftLimitSwitch;
    END_CASE;

    IF step <> prevStep THEN
        prevStep := step;
    ELSIF step > 0 THEN
        CASE step OF
            1: IF DownLimitSwitch THEN step := 0; prevStep := 0; END_IF;
            2: IF GripLimitSwitch THEN step := 0; prevStep := 0; END_IF;
            3: IF UpLimitSwitch THEN step := 0; prevStep := 0; END_IF;
            4: IF RightLimitSwitch THEN step := 0; prevStep := 0; END_IF;
            5: IF DownLimitSwitch THEN step := 0; prevStep := 0; END_IF;
            6: IF ReleaseLimitSwitch THEN step := 0; prevStep := 0; END_IF;
            7: IF UpLimitSwitch THEN step := 0; prevStep := 0; END_IF;
            8: IF LeftLimitSwitch THEN step := 0; prevStep := 0; END_IF;
        END_CASE;
    END_IF;

// Single cycle mode: Full sequence automatic, stop at end
ELSIF SingleCycleMode THEN
    IF startPressed THEN
        cycleActive := TRUE;
        prevStep := 0;
    END_IF;

    IF cycleActive THEN
        CASE step OF
            0: MoveDown := NOT DownLimitSwitch;
            1: ActivateGrip := NOT GripLimitSwitch;
            2: MoveUp := NOT UpLimitSwitch;
            3: MoveRight := NOT RightLimitSwitch;
            4: MoveDown := NOT DownLimitSwitch;
            5: ActivateRelease := NOT ReleaseLimitSwitch;
            6: MoveUp := NOT UpLimitSwitch;
            7: MoveLeft := NOT LeftLimitSwitch;
        END_CASE;

        IF step <> prevStep THEN
            prevStep := step;
        ELSIF step < 8 THEN
            CASE step OF
                0: IF DownLimitSwitch THEN step := 1; prevStep := 1; END_IF;
                1: IF GripLimitSwitch THEN step := 2; prevStep := 2; END_IF;
                2: IF UpLimitSwitch THEN step := 3; prevStep := 3; END_IF;
                3: IF RightLimitSwitch THEN step := 4; prevStep := 4; END_IF;
                4: IF DownLimitSwitch THEN step := 5; prevStep := 5; END_IF;
                5: IF ReleaseLimitSwitch THEN step := 6; prevStep := 6; END_IF;
                6: IF UpLimitSwitch THEN step := 7; prevStep := 7; END_IF;
                7: IF LeftLimitSwitch THEN step := 0; prevStep := 0; cycleActive := FALSE; END_IF;
            END_CASE;
        END_IF;
    END_IF;

// Continuous mode: Full sequence repeating
ELSIF ContinuousMode THEN
    IF startPressed THEN
        cycleActive := TRUE;
        prevStep := 0;
    END_IF;

    IF cycleActive THEN
        CASE step OF
            0: MoveDown := NOT DownLimitSwitch;
            1: ActivateGrip := NOT GripLimitSwitch;
            2: MoveUp := NOT UpLimitSwitch;
            3: MoveRight := NOT RightLimitSwitch;
            4: MoveDown := NOT DownLimitSwitch;
            5: ActivateRelease := NOT ReleaseLimitSwitch;
            6: MoveUp := NOT UpLimitSwitch;
            7: MoveLeft := NOT LeftLimitSwitch;
        END_CASE;

        IF step <> prevStep THEN
            prevStep := step;
        ELSIF step < 8 THEN
            CASE step OF
                0: IF DownLimitSwitch THEN step := 1; prevStep := 1; END_IF;
                1: IF GripLimitSwitch THEN step := 2; prevStep := 2; END_IF;
                2: IF UpLimitSwitch THEN step := 3; prevStep := 3; END_IF;
                3: IF RightLimitSwitch THEN step := 4; prevStep := 4; END_IF;
                4: IF DownLimitSwitch THEN step := 5; prevStep := 5; END_IF;
                5: IF ReleaseLimitSwitch THEN step := 6; prevStep := 6; END_IF;
                6: IF UpLimitSwitch THEN step := 7; prevStep := 7; END_IF;
                7: IF LeftLimitSwitch THEN step := 0; prevStep := 0; END_IF;
            END_CASE;
        END_IF;
    END_IF;

END_IF;
END_FUNCTION_BLOCK

(* ---- public-hard-05.raw_candidate_02.st ---- *)
FUNCTION_BLOCK MechanicalArmControl
VAR_INPUT
    ManualMode       : BOOL;
    SingleStepMode   : BOOL;
    SingleCycleMode  : BOOL;
    ContinuousMode   : BOOL;
    EmergencyStop    : BOOL;
    Start            : BOOL;
    DownButton       : BOOL;
    UpButton         : BOOL;
    LeftButton       : BOOL;
    RightButton      : BOOL;
    GripButton       : BOOL;
    ReleaseButton    : BOOL;
    DownLimitSwitch  : BOOL;
    UpLimitSwitch    : BOOL;
    LeftLimitSwitch  : BOOL;
    RightLimitSwitch : BOOL;
    GripLimitSwitch  : BOOL;
    ReleaseLimitSwitch : BOOL;
END_VAR

VAR_OUTPUT
    MoveDown       : BOOL;
    MoveUp         : BOOL;
    MoveLeft       : BOOL;
    MoveRight      : BOOL;
    ActivateGrip   : BOOL;
    ActivateRelease : BOOL;
END_VAR

VAR
    step         : UINT;
    prevStart    : BOOL;
    startPressed : BOOL;
    cycleActive  : BOOL;
END_VAR

// Reset all outputs first
MoveDown := FALSE;
MoveUp := FALSE;
MoveLeft := FALSE;
MoveRight := FALSE;
ActivateGrip := FALSE;
ActivateRelease := FALSE;

// Emergency stop: immediate halt
IF NOT EmergencyStop THEN
    step := 0;
    cycleActive := FALSE;
    prevStart := FALSE;
    RETURN;
END_IF;

// Rising edge detection for Start
startPressed := Start AND NOT prevStart;
prevStart := Start;

// Manual mode: Direct control via buttons
IF ManualMode THEN
    MoveDown := DownButton AND NOT DownLimitSwitch;
    MoveUp := UpButton AND NOT UpLimitSwitch;
    MoveLeft := LeftButton AND NOT LeftLimitSwitch;
    MoveRight := RightButton AND NOT RightLimitSwitch;
    ActivateGrip := GripButton;
    ActivateRelease := ReleaseButton;
    step := 0;
    cycleActive := FALSE;

// Single step mode: One action per Start press
ELSIF SingleStepMode THEN
    IF startPressed THEN
        step := step + 1;
        IF step > 8 THEN
            step := 1;
        END_IF;
    END_IF;

    // Execute current step
    CASE step OF
        1: MoveDown := NOT DownLimitSwitch;
        2: ActivateGrip := NOT GripLimitSwitch;
        3: MoveUp := NOT UpLimitSwitch;
        4: MoveRight := NOT RightLimitSwitch;
        5: MoveDown := NOT DownLimitSwitch;
        6: ActivateRelease := NOT ReleaseLimitSwitch;
        7: MoveUp := NOT UpLimitSwitch;
        8: MoveLeft := NOT LeftLimitSwitch;
    END_CASE;

    // Check completion and reset to wait for next Start
    CASE step OF
        1: IF DownLimitSwitch THEN step := 0; END_IF;
        2: IF GripLimitSwitch THEN step := 0; END_IF;
        3: IF UpLimitSwitch THEN step := 0; END_IF;
        4: IF RightLimitSwitch THEN step := 0; END_IF;
        5: IF DownLimitSwitch THEN step := 0; END_IF;
        6: IF ReleaseLimitSwitch THEN step := 0; END_IF;
        7: IF UpLimitSwitch THEN step := 0; END_IF;
        8: IF LeftLimitSwitch THEN step := 0; END_IF;
    END_CASE;

// Single cycle mode: Full sequence automatic, stop at end
ELSIF SingleCycleMode THEN
    IF startPressed THEN
        step := 0;
        cycleActive := TRUE;
    END_IF;

    IF cycleActive THEN
        CASE step OF
            0: MoveDown := NOT DownLimitSwitch;
            1: ActivateGrip := NOT GripLimitSwitch;
            2: MoveUp := NOT UpLimitSwitch;
            3: MoveRight := NOT RightLimitSwitch;
            4: MoveDown := NOT DownLimitSwitch;
            5: ActivateRelease := NOT ReleaseLimitSwitch;
            6: MoveUp := NOT UpLimitSwitch;
            7: MoveLeft := NOT LeftLimitSwitch;
        END_CASE;

        CASE step OF
            0: IF DownLimitSwitch THEN step := 1; END_IF;
            1: IF GripLimitSwitch THEN step := 2; END_IF;
            2: IF UpLimitSwitch THEN step := 3; END_IF;
            3: IF RightLimitSwitch THEN step := 4; END_IF;
            4: IF DownLimitSwitch THEN step := 5; END_IF;
            5: IF ReleaseLimitSwitch THEN step := 6; END_IF;
            6: IF UpLimitSwitch THEN step := 7; END_IF;
            7: IF LeftLimitSwitch THEN
                   step := 0;
                   cycleActive := FALSE;
               END_IF;
        END_CASE;
    END_IF;

// Continuous mode: Full sequence repeating
ELSIF ContinuousMode THEN
    IF startPressed THEN
        step := 0;
        cycleActive := TRUE;
    END_IF;

    IF cycleActive THEN
        CASE step OF
            0: MoveDown := NOT DownLimitSwitch;
            1: ActivateGrip := NOT GripLimitSwitch;
            2: MoveUp := NOT UpLimitSwitch;
            3: MoveRight := NOT RightLimitSwitch;
            4: MoveDown := NOT DownLimitSwitch;
            5: ActivateRelease := NOT ReleaseLimitSwitch;
            6: MoveUp := NOT UpLimitSwitch;
            7: MoveLeft := NOT LeftLimitSwitch;
        END_CASE;

        CASE step OF
            0: IF DownLimitSwitch THEN step := 1; END_IF;
            1: IF GripLimitSwitch THEN step := 2; END_IF;
            2: IF UpLimitSwitch THEN step := 3; END_IF;
            3: IF RightLimitSwitch THEN step := 4; END_IF;
            4: IF DownLimitSwitch THEN step := 5; END_IF;
            5: IF ReleaseLimitSwitch THEN step := 6; END_IF;
            6: IF UpLimitSwitch THEN step := 7; END_IF;
            7: IF LeftLimitSwitch THEN step := 0; END_IF;
        END_CASE;
    END_IF;

END_IF;
END_FUNCTION_BLOCK
